// TwinCAT 3 PLC project TcoAteqMeasurement
// Title: TcoAteqMeasurement
// Company: Vortex.Library
// ProjectVersion: 0.6.0.913
// ProgramVersion: 3.1.4023.0
// libraries:
//   Tc2_Standard, * (Beckhoff Automation GmbH)
//   Tc2_System, * (Beckhoff Automation GmbH)
//   Tc3_Module, * (Beckhoff Automation GmbH)
//   TcoIo, 0.6.0.913 (Vortex.Library)
//   TcoCore, 0.6.0.913 (Vortex.Library)
// project tree:
//   DUTs/G6/Enums/ eTcoAteqG6_AlarmCode_v_3_5_x.TcDUT, eTcoAteqG6_ParameterId_v_3_5_x.TcDUT, eTcoAteqG6_SpecialCycle_v_3_5_x.TcDUT, eTcoAteqG6_Step_v_3_5_x.TcDUT, eTcoAteqG6_TestType_v_3_5_x.TcDUT, eTcoAteqG6_Unit_v_3_5_x.TcDUT
//   DUTs/G6/ TcoAteqG6_CommandBits_v_3_5_x.TcDUT, TcoAteqG6_Config_v_3_5_x.TcDUT, TcoAteqG6_Control_v_3_5_x.TcDUT, TcoAteqG6_LastResult_v_3_5_x.TcDUT, TcoAteqG6_Measurement_v_3_5_x.TcDUT, TcoAteqG6_Parameter_v_3_5_x.TcDUT, TcoAteqG6_ParameterList_v_3_5_x.TcDUT, TcoAteqG6_ParameterQuery_v_3_5_x.TcDUT, TcoAteqG6_ParameterRequest_v_3_5_x.TcDUT, TcoAteqG6_ParameterSet_v_3_5_x.TcDUT, TcoAteqG6_State_v_3_5_x.TcDUT, TcoAteqG6_Status_v_3_5_x.TcDUT, TcoAteqG6_StatusBits_v_3_5_x.TcDUT
//   / PlcTask.TcTTO
//   POUs/Functions/G6/ TcoAteqG6_AddParameterToRequest_v_3_5_x.TcPOU, TcoAteqG6_BuildPresetRequest_v_3_5_x.TcPOU, TcoAteqG6_ClearLastResult_v_3_5_x.TcPOU, TcoAteqG6_ClearMeasurement_v_3_5_x.TcPOU, TcoAteqG6_ClearParameterList_v_3_5_x.TcPOU, TcoAteqG6_ClearParameterRequest_v_3_5_x.TcPOU, TcoAteqG6_DecodeCommandBits_v_3_5_x.TcPOU, TcoAteqG6_DecodeLastResult_v_3_5_x.TcPOU, TcoAteqG6_DecodeMeasurement_v_3_5_x.TcPOU, TcoAteqG6_DecodeParameterList_v_3_5_x.TcPOU, TcoAteqG6_DecodeState_v_3_5_x.TcPOU, TcoAteqG6_DecodeStatusBits_v_3_5_x.TcPOU, TcoAteqG6_EncodeControl_v_3_5_x.TcPOU, TcoAteqG6_GetDint_v_3_5_x.TcPOU, TcoAteqG6_GetInt_v_3_5_x.TcPOU, TcoAteqG6_GetWord_v_3_5_x.TcPOU, TcoAteqG6_IsParameterRequestValid_v_3_5_x.TcPOU, TcoAteqG6_MapPresetParameters_v_3_5_x.TcPOU, TcoAteqG6_QueryParameter_v_3_5_x.TcPOU, TcoAteqG6_SetDint_v_3_5_x.TcPOU, TcoAteqG6_SetWord_v_3_5_x.TcPOU, TcoAteqG6_SpecialCycleToByte_v_3_5_x.TcPOU, TcoAteqG6_ToAlarmCode_v_3_5_x.TcPOU, TcoAteqG6_ToEngineering_v_3_5_x.TcPOU, TcoAteqG6_ToStep_v_3_5_x.TcPOU, TcoAteqG6_ToTestType_v_3_5_x.TcPOU, TcoAteqG6_ToUnit_v_3_5_x.TcPOU, TcoAteqG6_TryGetParameterRaw_v_3_5_x.TcPOU
//   POUs/ MAIN.TcPOU
//   POUs/Prototypes/G6/IO/ TcoAteqG6_Inputs_v_3_5_x.TcDUT, TcoAteqG6_Outputs_v_3_5_x.TcDUT, TcoAteqG6Pn_IO_v_3_5_x.TcDUT
//   POUs/Prototypes/G6/ TcoAteqG6Pn_v_3_5_x.TcPOU
//   POUs/Prototypes/MeasurementTasks/G6_v_3_5_x/ TcoAteqG6_ReadLastResultTask_v_3_5_x.TcPOU, TcoAteqG6_ReadParametersTask_v_3_5_x.TcPOU, TcoAteqG6_ResetTask_v_3_5_x.TcPOU, TcoAteqG6_SelectProgramTask_v_3_5_x.TcPOU, TcoAteqG6_SpecialCycleTask_v_3_5_x.TcPOU, TcoAteqG6_StartCycleTask_v_3_5_x.TcPOU, TcoAteqG6Task_v_3_5_x.TcPOU
// real-time tasks:
//   TASK PlcTask: cycle T#10ms, priority 20, ADS port 350
//   TASK PlcTask1: cycle T#10ms, priority 21, ADS port 351

CONFIGURATION TcoAteqMeasurement
    RESOURCE PLC ON TwinCAT3
        TASK PlcTask(INTERVAL := T#10ms, PRIORITY := 20);
        PROGRAM MAIN WITH PlcTask : MAIN;
    END_RESOURCE
END_CONFIGURATION

// ---- DUTs/G6/Enums/eTcoAteqG6_AlarmCode_v_3_5_x.TcDUT
(*~
	<docu>
		<summary>
			Alarm code of the last result (exchange zone 26h). Codes that are not listed decode to Unknown.
		</summary>
	</docu>
~*)
{attribute 'qualified_only'}
{attribute 'strict'}
TYPE eTcoAteqG6_AlarmCode_v_3_5_x :
(
	Unknown := -1,
	NoAlarm := 0,
	PressureSwitchTooHigh := 1,
	PressureSwitchTooLow := 2,
	LargeLeakOnTest := 3,
	LargeLeakOnReference := 4,
	SensorOutOfOrder := 7,
	PressureTooHigh := 43,
	PressureTooLow := 44,
	PiezoSensorOutOfOrder := 45,
	DumpError := 46,
	CalibrationDrift := 47,
	AtmosphericPressureError := 73,
	TemperatureError := 74
) INT;
END_TYPE

// ---- DUTs/G6/Enums/eTcoAteqG6_ParameterId_v_3_5_x.TcDUT
(*~
	<docu>
		<summary>
			Parameter identifiers of the "Read parameters" command (manual pp. 43-46). Every value is exchanged as LONG x1000; times in seconds, levels in the instrument units, selections as code x1000.
		</summary>
	</docu>
~*)
{attribute 'qualified_only'}
{attribute 'strict'}
TYPE eTcoAteqG6_ParameterId_v_3_5_x :
(
	None := 0,
	FillTime := 1,
	StabTime := 2,
	TestTime := 3,
	PreFillTime := 6,
	DumpTime := 9,
	CouplingTimeA := 10,
	CouplingTimeB := 11,
	PartVolume := 20,
	TestType := 21,
	InterCycleTime := 29,
	ResultHoldTime := 48,
	MinFill := 50,
	MaxFill := 51,
	PressureUnit := 53,
	TestFail := 60,
	TestRework := 61,
	RefFail := 62,
	RefRework := 63,
	SetFill := 66,
	DiffAutoResetTime := 80,
	FillMode := 103,
	ExternalDumpType := 110,
	Input7Function := 112,
	Language := 123,
	MaxPreFill := 126,
	FlowUnit := 127,
	CalibrationLeakRate := 128,
	Filter := 148,
	UnitType := 149,
	BarGraphMaxReject := 158,
	VolumeUnit := 161,
	NextProgram := 164,
	PiezoAutoZeroCycles := 165,
	PiezoAutoZeroMinutes := 166,
	DelayExt1 := 249,
	DelayExt2 := 250,
	DelayExt3 := 251,
	DelayExt4 := 252,
	DelayExt5 := 253,
	DelayExt6 := 254,
	DelayInt2 := 255,
	DelayInt1 := 256,
	DelayAux1 := 257,
	DelayAux2 := 258,
	DelayAux3 := 259,
	DelayAux4 := 260,
	TimeExt1 := 261,
	TimeExt2 := 262,
	TimeExt3 := 263,
	TimeExt4 := 264,
	TimeExt5 := 265,
	TimeExt6 := 266,
	TimeInt2 := 267,
	TimeInt1 := 268,
	TimeAux1 := 269,
	TimeAux2 := 270,
	TimeAux3 := 271,
	TimeAux4 := 272,
	PressureFilter := 274,
	CapillaryRange := 281,
	BarCodeFirstChar := 287,
	BarCodeCharCount := 288,
	BarCodeProgram := 289,
	GeneralPressureUnit := 353,
	LinePressureMin := 354,
	DisplayMode := 364,
	Input8Function := 375,
	Input9Function := 376,
	UsbMode := 379,
	SaveOn := 412,
	AccessMode := 413,
	Year := 414,
	Month := 415,
	Day := 416,
	Hour := 417,
	Minute := 418,
	Second := 419,
	LearningCycles := 459,
	LearningInterCycleTime := 460,
	LearningMaxOffset := 461,
	LearningFlowMaster := 462,
	LearningPressureMaster := 463,
	LearningMinVolume := 464,
	LearningMaxVolume := 465,
	LearningOffset := 486
) UINT;
END_TYPE

// ---- DUTs/G6/Enums/eTcoAteqG6_SpecialCycle_v_3_5_x.TcDUT
(*~
	<docu>
		<summary>
			Special cycle table (manual p. 58). Ids 25..31 require the "Service" special-cycle function to be enabled on the instrument.
		</summary>
	</docu>
~*)
{attribute 'qualified_only'}
{attribute 'strict'}
TYPE eTcoAteqG6_SpecialCycle_v_3_5_x :
(
	None := 0,
	AtrLearning := 1,
	CustomUnitLearn := 4,
	CustomUnitCheck := 5,
	PiezoAutoZero := 9,
	RegulatorAdjust := 13,
	CapillaryTemperatureCheck := 25,
	TemperatureCheck := 26,
	AtmPressureCheck := 27,
	P1SensorCheck := 28,
	Flow1Check := 29,
	Flow2Check := 30,
	LinePressureSensorCheck := 31
) INT;
END_TYPE

// ---- DUTs/G6/Enums/eTcoAteqG6_Step_v_3_5_x.TcDUT
(*~
	<docu>
		<summary>
			Current test step (input 0Eh). None = FFFFh on the bus (no cycle running).
		</summary>
	</docu>
~*)
{attribute 'qualified_only'}
{attribute 'strict'}
TYPE eTcoAteqG6_Step_v_3_5_x :
(
	Unknown := -2,
	None := -1,
	PreFill := 0,
	Fill := 1,
	ZeroDiff := 2,
	Stabilization := 3,
	Test := 4,
	Dump := 5
) INT;
END_TYPE

// ---- DUTs/G6/Enums/eTcoAteqG6_TestType_v_3_5_x.TcDUT
(*~
	<docu>
		<summary>
			Test type parameter (id 21).
		</summary>
	</docu>
~*)
{attribute 'qualified_only'}
{attribute 'strict'}
TYPE eTcoAteqG6_TestType_v_3_5_x :
(
	Unknown := -1,
	Invalid := 0,
	Direct := 1,
	Operator := 2
) INT;
END_TYPE

// ---- DUTs/G6/Enums/eTcoAteqG6_Unit_v_3_5_x.TcDUT
(*~
	<docu>
		<summary>
			Unit table (manual p. 48). On the bus a unit is a LONG holding the unit code; the enum value is that code divided by 1000 (14000 = mbar).
		</summary>
	</docu>
~*)
{attribute 'qualified_only'}
{attribute 'strict'}
TYPE eTcoAteqG6_Unit_v_3_5_x :
(
	Unknown := -1,
	cm3_s := 0,
	cm3_min := 1,
	cm3_h := 2,
	Pa := 6,
	bar := 11,
	kPa := 12,
	PSI := 13,
	mbar := 14,
	MPa := 15,
	l_h := 30,
	inch3_s := 46,
	inch3_min := 47,
	inch3_h := 48,
	ft3_h := 49,
	ml_s := 50,
	ml_min := 51,
	ml_h := 52,
	mm3 := 55,
	cm3 := 56,
	ml := 61,
	l := 62,
	inch3 := 63,
	ft3 := 64,
	SCCM := 84,
	Points := 92
) INT;
END_TYPE

// ---- DUTs/G6/TcoAteqG6_CommandBits_v_3_5_x.TcDUT
(*~
	<docu>
		<summary>
			Bit view of a command, echo or error word (bit 0 = Reset ... bit 15 = Read last result).
		</summary>
	</docu>
~*)
TYPE TcoAteqG6_CommandBits_v_3_5_x :
STRUCT
	{attribute addProperty Name "<#Raw#>"}
	Raw : WORD;
	{attribute addProperty Name "<#Reset#>"}
	Reset : BOOL;
	{attribute addProperty Name "<#Start#>"}
	Start : BOOL;
	{attribute addProperty Name "<#Special cycle#>"}
	SpecialCycle : BOOL;
	{attribute addProperty Name "<#Program selection#>"}
	ProgramSelection : BOOL;
	{attribute addProperty Name "<#Read FIFO results#>"}
	ReadFifo : BOOL;
	{attribute addProperty Name "<#Read parameters#>"}
	ReadParameters : BOOL;
	{attribute addProperty Name "<#Write parameters#>"}
	WriteParameters : BOOL;
	{attribute addProperty Name "<#Reset FIFO results#>"}
	ResetFifo : BOOL;
	{attribute addProperty Name "<#Read instrument configuration#>"}
	ReadInstrumentConfiguration : BOOL;
	{attribute addProperty Name "<#Read configuration bits#>"}
	ReadConfigurationBits : BOOL;
	{attribute addProperty Name "<#Read function bits#>"}
	ReadFunctionBits : BOOL;
	{attribute addProperty Name "<#Write configuration bits#>"}
	WriteConfigurationBits : BOOL;
	{attribute addProperty Name "<#Write function bits#>"}
	WriteFunctionBits : BOOL;
	{attribute addProperty Name "<#Read program name#>"}
	ReadProgramName : BOOL;
	{attribute addProperty Name "<#Write program name#>"}
	WriteProgramName : BOOL;
	{attribute addProperty Name "<#Read last result#>"}
	ReadLastResult : BOOL;
END_STRUCT
END_TYPE

// ---- DUTs/G6/TcoAteqG6_Config_v_3_5_x.TcDUT
(*~
	<docu>
		<summary>
			Configuration of TcoAteqG6Pn_v_3_5_x. CommandTimeout / CycleTimeout of 0 fall back to 5 s / 60 s.
		</summary>
	</docu>
~*)
TYPE TcoAteqG6_Config_v_3_5_x :
STRUCT
	{attribute addProperty Name "<#Info time#>"}
	InfoTime : TIME := T#2S;
	{attribute addProperty Name "<#Task timeout (0 = off)#>"}
	ErrorTime : TIME := T#0S;
	{attribute addProperty Name "<#Command handshake timeout (per step)#>"}
	CommandTimeout : TIME := T#5S;
	{attribute addProperty Name "<#Test cycle timeout#>"}
	CycleTimeout : TIME := T#60S;
END_STRUCT
END_TYPE

// ---- DUTs/G6/TcoAteqG6_Control_v_3_5_x.TcDUT
(*~
	<docu>
		<summary>
			Output data: 00h command word, 06h program number (0-based on the bus), 08h special cycle id, 09h special cycle instruction, 20h parameter request. The whole output image is rewritten every cycle.
		</summary>
	</docu>
~*)
TYPE TcoAteqG6_Control_v_3_5_x :
STRUCT
	{attribute addProperty Name "<#Command word#>"}
	Command : WORD;
	{attribute addProperty Name "<#Command bits#>"}
	CommandBits : TcoAteqG6_CommandBits_v_3_5_x;
	{attribute addProperty Name "<#Program number (as displayed, 1-128)#>"}
	ProgramNumber : INT;
	{attribute addProperty Name "<#Special cycle#>"}
	SpecialCycle : eTcoAteqG6_SpecialCycle_v_3_5_x;
	{attribute addProperty Name "<#Special cycle instruction#>"}
	SpecialCycleInstruction : BYTE;
	{attribute addProperty Name "<#Parameter request#>"}
	ParameterRequest : TcoAteqG6_ParameterRequest_v_3_5_x;
	{attribute addProperty Name "<#Selected parameter#>"}
	QueryParameter : eTcoAteqG6_ParameterId_v_3_5_x;
END_STRUCT
END_TYPE

// ---- DUTs/G6/TcoAteqG6_LastResult_v_3_5_x.TcDUT
(*~
	<docu>
		<summary>
			Last result, decoded from the exchange zone (20h..37h) after the "Read last result" command. Valid = no alarm.
		</summary>
	</docu>
~*)
TYPE TcoAteqG6_LastResult_v_3_5_x :
STRUCT
	{attribute addProperty Name "<#Valid#>"}
	Valid : BOOL;
	{attribute addProperty Name "<#Program#>"}
	ProgramNo : INT;
	{attribute addProperty Name "<#Test type (raw)#>"}
	TestTypeRaw : INT;
	{attribute addProperty Name "<#Pass#>"}
	Pass : BOOL;
	{attribute addProperty Name "<#Fail test part (maximum flow reject)#>"}
	FailTest : BOOL;
	{attribute addProperty Name "<#Fail reference part (minimum flow reject)#>"}
	FailReference : BOOL;
	{attribute addProperty Name "<#Alarm#>"}
	Alarm : BOOL;
	{attribute addProperty Name "<#Pressure error (unverified)#>"}
	PressureError : BOOL;
	{attribute addProperty Name "<#Part recoverable (unverified)#>"}
	Recoverable : BOOL;
	{attribute addProperty Name "<#Calibration error (unverified)#>"}
	CalibrationError : BOOL;
	{attribute addProperty Name "<#Calibration check error (unverified)#>"}
	CalibrationCheckError : BOOL;
	{attribute addProperty Name "<#ATR fault (unverified)#>"}
	AtrFault : BOOL;
	{attribute addProperty Name "<#Relay image (raw)#>"}
	RelayImageRaw : WORD;
	{attribute addProperty Name "<#Alarm code#>"}
	AlarmCode : eTcoAteqG6_AlarmCode_v_3_5_x;
	{attribute addProperty Name "<#Alarm code (raw)#>"}
	AlarmCodeRaw : INT;
	{attribute addProperty Name "<#Measurement#>"}
	Measurement : TcoAteqG6_Measurement_v_3_5_x;
END_STRUCT
END_TYPE

// ---- DUTs/G6/TcoAteqG6_Measurement_v_3_5_x.TcDUT
(*~
	<docu>
		<summary>
			Pressure and flow with their units: four LONGs (value x1000, unit code).
		</summary>
	</docu>
~*)
TYPE TcoAteqG6_Measurement_v_3_5_x :
STRUCT
	{attribute addProperty Name "<#Pressure#>"}
	Pressure : REAL;
	{attribute addProperty Name "<#Pressure unit#>"}
	PressureUnit : eTcoAteqG6_Unit_v_3_5_x := eTcoAteqG6_Unit_v_3_5_x.Unknown;
	{attribute addProperty Name "<#Flow / leak#>"}
	Flow : REAL;
	{attribute addProperty Name "<#Flow unit#>"}
	FlowUnit : eTcoAteqG6_Unit_v_3_5_x := eTcoAteqG6_Unit_v_3_5_x.Unknown;
	{attribute addProperty Name "<#Pressure (raw x1000)#>"}
	PressureRaw : DINT;
	{attribute addProperty Name "<#Pressure unit code (raw)#>"}
	PressureUnitRaw : DINT;
	{attribute addProperty Name "<#Flow (raw x1000)#>"}
	FlowRaw : DINT;
	{attribute addProperty Name "<#Flow unit code (raw)#>"}
	FlowUnitRaw : DINT;
END_STRUCT
END_TYPE

// ---- DUTs/G6/TcoAteqG6_Parameter_v_3_5_x.TcDUT
(*~
	<docu>
		<summary>
			One parameter of the "Read parameters" response.
		</summary>
	</docu>
~*)
TYPE TcoAteqG6_Parameter_v_3_5_x :
STRUCT
	{attribute addProperty Name "<#Identifier#>"}
	Id : UINT;
	{attribute addProperty Name "<#Value#>"}
	Value : REAL;
	{attribute addProperty Name "<#Value (raw x1000)#>"}
	Raw : DINT;
END_STRUCT
END_TYPE

// ---- DUTs/G6/TcoAteqG6_ParameterList_v_3_5_x.TcDUT
(*~
	<docu>
		<summary>
			Response of the "Read parameters" command: from input 20h one identifier WORD + value LONG x1000 per parameter.
		</summary>
	</docu>
~*)
TYPE TcoAteqG6_ParameterList_v_3_5_x :
STRUCT
	{attribute addProperty Name "<#Number of parameters read#>"}
	Count : INT;
	{attribute addProperty Name "<#Parameters#>"}
	Items : ARRAY[0..34] OF TcoAteqG6_Parameter_v_3_5_x;
END_STRUCT
END_TYPE

// ---- DUTs/G6/TcoAteqG6_ParameterQuery_v_3_5_x.TcDUT
(*~
	<docu>
		<summary>
			Value of the selected parameter (Control.QueryParameter), looked up after every "Read parameters".
		</summary>
	</docu>
~*)
TYPE TcoAteqG6_ParameterQuery_v_3_5_x :
STRUCT
	{attribute addProperty Name "<#Parameter#>"}
	Parameter : eTcoAteqG6_ParameterId_v_3_5_x;
	{attribute addProperty Name "<#Found#>"}
	Found : BOOL;
	{attribute addProperty Name "<#Value#>"}
	Value : REAL;
	{attribute addProperty Name "<#Value (raw x1000)#>"}
	Raw : DINT;
END_STRUCT
END_TYPE

// ---- DUTs/G6/TcoAteqG6_ParameterRequest_v_3_5_x.TcDUT
(*~
	<docu>
		<summary>
			Request of the "Read parameters" command (output 20h: count, then up to 35 identifiers).
		</summary>
	</docu>
~*)
TYPE TcoAteqG6_ParameterRequest_v_3_5_x :
STRUCT
	{attribute addProperty Name "<#Number of parameters (1-35)#>"}
	Count : INT;
	{attribute addProperty Name "<#Identifiers#>"}
	Ids : ARRAY[0..34] OF UINT;
END_STRUCT
END_TYPE

// ---- DUTs/G6/TcoAteqG6_ParameterSet_v_3_5_x.TcDUT
(*~
	<docu>
		<summary>
			Typed view of the commonly used program parameters (manual p. 43), filled by ReadPresetParameters.
		</summary>
	</docu>
~*)
TYPE TcoAteqG6_ParameterSet_v_3_5_x :
STRUCT
	{attribute addProperty Name "<#Fill time [s]#>"}
	FillTime : REAL;
	{attribute addProperty Name "<#Stabilization time [s]#>"}
	StabTime : REAL;
	{attribute addProperty Name "<#Test time [s]#>"}
	TestTime : REAL;
	{attribute addProperty Name "<#Dump time [s]#>"}
	DumpTime : REAL;
	{attribute addProperty Name "<#Test type#>"}
	TestType : eTcoAteqG6_TestType_v_3_5_x;
	{attribute addProperty Name "<#Minimum fill pressure#>"}
	MinFill : REAL;
	{attribute addProperty Name "<#Maximum fill pressure#>"}
	MaxFill : REAL;
	{attribute addProperty Name "<#Pressure unit#>"}
	PressureUnit : eTcoAteqG6_Unit_v_3_5_x := eTcoAteqG6_Unit_v_3_5_x.Unknown;
	{attribute addProperty Name "<#Test part reject level#>"}
	TestFail : REAL;
	{attribute addProperty Name "<#Reference part reject level#>"}
	RefFail : REAL;
	{attribute addProperty Name "<#Fill set point#>"}
	SetFill : REAL;
END_STRUCT
END_TYPE

// ---- DUTs/G6/TcoAteqG6_State_v_3_5_x.TcDUT
(*~
	<docu>
		<summary>
			Decoded input image: 00h echo, 02h error word (FFFFh = command running), 06h program (0-based on the bus), 08h results in FIFO, 0Ah test type, 0Ch status bits, 0Eh step, 10h..1Fh real-time pressure/flow.
		</summary>
	</docu>
~*)
TYPE TcoAteqG6_State_v_3_5_x :
STRUCT
	{attribute addProperty Name "<#Command echo#>"}
	Echo : TcoAteqG6_CommandBits_v_3_5_x;
	{attribute addProperty Name "<#Command error#>"}
	Error : TcoAteqG6_CommandBits_v_3_5_x;
	{attribute addProperty Name "<#Command running#>"}
	CommandRunning : BOOL;
	{attribute addProperty Name "<#Current program#>"}
	CurrentProgram : INT;
	{attribute addProperty Name "<#Results in FIFO#>"}
	ResultsInFifo : INT;
	{attribute addProperty Name "<#Test type (raw)#>"}
	TestTypeRaw : INT;
	{attribute addProperty Name "<#Status#>"}
	StatusBits : TcoAteqG6_StatusBits_v_3_5_x;
	{attribute addProperty Name "<#Step#>"}
	Step : eTcoAteqG6_Step_v_3_5_x := eTcoAteqG6_Step_v_3_5_x.None;
	{attribute addProperty Name "<#Step (raw)#>"}
	StepRaw : INT;
	{attribute addProperty Name "<#Real time#>"}
	RealTime : TcoAteqG6_Measurement_v_3_5_x;
END_STRUCT
END_TYPE

// ---- DUTs/G6/TcoAteqG6_Status_v_3_5_x.TcDUT
(*~
	<docu>
		<summary>
			Status of TcoAteqG6Pn_v_3_5_x.
		</summary>
	</docu>
~*)
TYPE TcoAteqG6_Status_v_3_5_x :
STRUCT
	{attribute addProperty Name "<#Action#>"}
	ActionDescription : STRING(100);
	{attribute addProperty Name "<#Ready#>"}
	Ready : BOOL;
	{attribute addProperty Name "<#Last part passed#>"}
	LastPass : BOOL;
	{attribute addProperty Name "<#Last command error word#>"}
	LastCommandError : WORD;
	{attribute addProperty Name "<#Instrument#>"}
	State : TcoAteqG6_State_v_3_5_x;
	{attribute addProperty Name "<#Last result#>"}
	LastResult : TcoAteqG6_LastResult_v_3_5_x;
	{attribute addProperty Name "<#Parameters#>"}
	Parameters : TcoAteqG6_ParameterList_v_3_5_x;
	{attribute addProperty Name "<#Preset parameters#>"}
	ParameterSet : TcoAteqG6_ParameterSet_v_3_5_x;
	{attribute addProperty Name "<#Selected parameter#>"}
	ParameterQuery : TcoAteqG6_ParameterQuery_v_3_5_x;
END_STRUCT
END_TYPE

// ---- DUTs/G6/TcoAteqG6_StatusBits_v_3_5_x.TcDUT
(*~
	<docu>
		<summary>
			Status word of the instrument (input 0Ch). Bits 8 and 10..14 are not used.
		</summary>
	</docu>
~*)
TYPE TcoAteqG6_StatusBits_v_3_5_x :
STRUCT
	{attribute addProperty Name "<#Raw#>"}
	Raw : WORD;
	{attribute addProperty Name "<#Pass#>"}
	Pass : BOOL;
	{attribute addProperty Name "<#Fail test part#>"}
	FailTest : BOOL;
	{attribute addProperty Name "<#Fail reference part#>"}
	FailReference : BOOL;
	{attribute addProperty Name "<#Alarm#>"}
	Alarm : BOOL;
	{attribute addProperty Name "<#Pressure error#>"}
	PressureError : BOOL;
	{attribute addProperty Name "<#Cycle end#>"}
	CycleEnd : BOOL;
	{attribute addProperty Name "<#Part recoverable#>"}
	Recoverable : BOOL;
	{attribute addProperty Name "<#Calibration error or drift#>"}
	CalibrationError : BOOL;
	{attribute addProperty Name "<#ATR error or drift#>"}
	AtrError : BOOL;
	{attribute addProperty Name "<#Key presence#>"}
	KeyPresence : BOOL;
END_STRUCT
END_TYPE

// ---- POUs/Prototypes/G6/IO/TcoAteqG6_Inputs_v_3_5_x.TcDUT
TYPE TcoAteqG6_Inputs_v_3_5_x :
STRUCT
	{attribute addProperty Name "<#Input module 1 (slot 1, 00h..3Fh)#>"}
	In1 AT %I* : ARRAY[0..63] OF BYTE;
	{attribute addProperty Name "<#Input module 2 (slot 2, 40h..7Fh)#>"}
	In2 AT %I* : ARRAY[0..63] OF BYTE;
	{attribute addProperty Name "<#Input module 3 (slot 3, 80h..BFh)#>"}
	In3 AT %I* : ARRAY[0..63] OF BYTE;
	{attribute addProperty Name "<#Input module 4 (slot 4, C0h..FFh)#>"}
	In4 AT %I* : ARRAY[0..63] OF BYTE;
END_STRUCT
END_TYPE

// ---- POUs/Prototypes/G6/IO/TcoAteqG6_Outputs_v_3_5_x.TcDUT
TYPE TcoAteqG6_Outputs_v_3_5_x :
STRUCT
	{attribute addProperty Name "<#Output module 1 (slot 5, 00h..3Fh)#>"}
	Out1 AT %Q* : ARRAY[0..63] OF BYTE;
	{attribute addProperty Name "<#Output module 2 (slot 6, 40h..7Fh)#>"}
	Out2 AT %Q* : ARRAY[0..63] OF BYTE;
	{attribute addProperty Name "<#Output module 3 (slot 7, 80h..BFh)#>"}
	Out3 AT %Q* : ARRAY[0..63] OF BYTE;
	{attribute addProperty Name "<#Output module 4 (slot 8, C0h..FFh)#>"}
	Out4 AT %Q* : ARRAY[0..63] OF BYTE;
END_STRUCT
END_TYPE

// ---- POUs/Prototypes/G6/IO/TcoAteqG6Pn_IO_v_3_5_x.TcDUT
TYPE TcoAteqG6Pn_IO_v_3_5_x :
STRUCT
	PnIoBoxState AT %I*	:	UINT;
	PnIoBoxDiag AT %I*	:	UINT;
	PnIoBoxCtrl AT %Q*	:	UINT;
	{attribute addProperty Name "<#IN#>"}
	In : TcoAteqG6_Inputs_v_3_5_x;
	{attribute addProperty Name "<#OUT#>"}
	Out : TcoAteqG6_Outputs_v_3_5_x;
END_STRUCT
END_TYPE

// ---- POUs/MAIN.TcPOU
PROGRAM MAIN
VAR
END_VAR

END_PROGRAM

// ---- POUs/Functions/G6/TcoAteqG6_AddParameterToRequest_v_3_5_x.TcPOU
(*~
	<docu>
		<summary>
			Appends a parameter identifier to the request. Returns FALSE when the request is full (35).
		</summary>
	</docu>
~*)
FUNCTION TcoAteqG6_AddParameterToRequest_v_3_5_x : BOOL
VAR_INPUT
	inParameter : eTcoAteqG6_ParameterId_v_3_5_x;
END_VAR
VAR_IN_OUT
	inoRequest : TcoAteqG6_ParameterRequest_v_3_5_x;
END_VAR

IF inoRequest.Count < 0 OR inoRequest.Count >= 35 THEN
	RETURN;
END_IF
inoRequest.Ids[inoRequest.Count] := TO_UINT(inParameter);
inoRequest.Count := inoRequest.Count + 1;
TcoAteqG6_AddParameterToRequest_v_3_5_x := TRUE;

END_FUNCTION

// ---- POUs/Functions/G6/TcoAteqG6_BuildPresetRequest_v_3_5_x.TcPOU
(*~
	<docu>
		<summary>
			Fills the request with the 11 identifiers of the preset parameter set.
		</summary>
	</docu>
~*)
FUNCTION TcoAteqG6_BuildPresetRequest_v_3_5_x : BOOL
VAR_IN_OUT
	inoRequest : TcoAteqG6_ParameterRequest_v_3_5_x;
END_VAR

TcoAteqG6_ClearParameterRequest_v_3_5_x(inoRequest := inoRequest);
TcoAteqG6_AddParameterToRequest_v_3_5_x(inParameter := eTcoAteqG6_ParameterId_v_3_5_x.FillTime, inoRequest := inoRequest);
TcoAteqG6_AddParameterToRequest_v_3_5_x(inParameter := eTcoAteqG6_ParameterId_v_3_5_x.StabTime, inoRequest := inoRequest);
TcoAteqG6_AddParameterToRequest_v_3_5_x(inParameter := eTcoAteqG6_ParameterId_v_3_5_x.TestTime, inoRequest := inoRequest);
TcoAteqG6_AddParameterToRequest_v_3_5_x(inParameter := eTcoAteqG6_ParameterId_v_3_5_x.DumpTime, inoRequest := inoRequest);
TcoAteqG6_AddParameterToRequest_v_3_5_x(inParameter := eTcoAteqG6_ParameterId_v_3_5_x.TestType, inoRequest := inoRequest);
TcoAteqG6_AddParameterToRequest_v_3_5_x(inParameter := eTcoAteqG6_ParameterId_v_3_5_x.MinFill, inoRequest := inoRequest);
TcoAteqG6_AddParameterToRequest_v_3_5_x(inParameter := eTcoAteqG6_ParameterId_v_3_5_x.MaxFill, inoRequest := inoRequest);
TcoAteqG6_AddParameterToRequest_v_3_5_x(inParameter := eTcoAteqG6_ParameterId_v_3_5_x.PressureUnit, inoRequest := inoRequest);
TcoAteqG6_AddParameterToRequest_v_3_5_x(inParameter := eTcoAteqG6_ParameterId_v_3_5_x.TestFail, inoRequest := inoRequest);
TcoAteqG6_AddParameterToRequest_v_3_5_x(inParameter := eTcoAteqG6_ParameterId_v_3_5_x.RefFail, inoRequest := inoRequest);
TcoAteqG6_AddParameterToRequest_v_3_5_x(inParameter := eTcoAteqG6_ParameterId_v_3_5_x.SetFill, inoRequest := inoRequest);
TcoAteqG6_BuildPresetRequest_v_3_5_x := TRUE;

END_FUNCTION

// ---- POUs/Functions/G6/TcoAteqG6_ClearParameterRequest_v_3_5_x.TcPOU
(*~
	<docu>
		<summary>
			Clears a parameter request.
		</summary>
	</docu>
~*)
FUNCTION TcoAteqG6_ClearParameterRequest_v_3_5_x : BOOL
VAR_IN_OUT
	inoRequest : TcoAteqG6_ParameterRequest_v_3_5_x;
END_VAR
VAR
	i : INT;
END_VAR

inoRequest.Count := 0;
FOR i := 0 TO 34 DO
	inoRequest.Ids[i] := 0;
END_FOR
TcoAteqG6_ClearParameterRequest_v_3_5_x := TRUE;

END_FUNCTION

// ---- POUs/Functions/G6/TcoAteqG6_ClearLastResult_v_3_5_x.TcPOU
(*~
	<docu>
		<summary>
			Clears the last result (Valid = FALSE).
		</summary>
	</docu>
~*)
FUNCTION TcoAteqG6_ClearLastResult_v_3_5_x : BOOL
VAR_IN_OUT
	inoResult : TcoAteqG6_LastResult_v_3_5_x;
END_VAR

inoResult.Valid := FALSE;
inoResult.ProgramNo := 0;
inoResult.TestTypeRaw := 0;
inoResult.Pass := FALSE;
inoResult.FailTest := FALSE;
inoResult.FailReference := FALSE;
inoResult.Alarm := FALSE;
inoResult.PressureError := FALSE;
inoResult.Recoverable := FALSE;
inoResult.CalibrationError := FALSE;
inoResult.CalibrationCheckError := FALSE;
inoResult.AtrFault := FALSE;
inoResult.RelayImageRaw := 0;
inoResult.AlarmCode := eTcoAteqG6_AlarmCode_v_3_5_x.NoAlarm;
inoResult.AlarmCodeRaw := 0;
TcoAteqG6_ClearMeasurement_v_3_5_x(inoMeasurement := inoResult.Measurement);
TcoAteqG6_ClearLastResult_v_3_5_x := TRUE;

END_FUNCTION

// ---- POUs/Functions/G6/TcoAteqG6_ClearMeasurement_v_3_5_x.TcPOU
(*~
	<docu>
		<summary>
			Clears a measurement.
		</summary>
	</docu>
~*)
FUNCTION TcoAteqG6_ClearMeasurement_v_3_5_x : BOOL
VAR_IN_OUT
	inoMeasurement : TcoAteqG6_Measurement_v_3_5_x;
END_VAR

inoMeasurement.Pressure := 0.0;
inoMeasurement.PressureUnit := eTcoAteqG6_Unit_v_3_5_x.Unknown;
inoMeasurement.Flow := 0.0;
inoMeasurement.FlowUnit := eTcoAteqG6_Unit_v_3_5_x.Unknown;
inoMeasurement.PressureRaw := 0;
inoMeasurement.PressureUnitRaw := 0;
inoMeasurement.FlowRaw := 0;
inoMeasurement.FlowUnitRaw := 0;
TcoAteqG6_ClearMeasurement_v_3_5_x := TRUE;

END_FUNCTION

// ---- POUs/Functions/G6/TcoAteqG6_ClearParameterList_v_3_5_x.TcPOU
(*~
	<docu>
		<summary>
			Clears a parameter list.
		</summary>
	</docu>
~*)
FUNCTION TcoAteqG6_ClearParameterList_v_3_5_x : BOOL
VAR_IN_OUT
	inoList : TcoAteqG6_ParameterList_v_3_5_x;
END_VAR
VAR
	i : INT;
END_VAR

inoList.Count := 0;
FOR i := 0 TO 34 DO
	inoList.Items[i].Id := 0;
	inoList.Items[i].Raw := 0;
	inoList.Items[i].Value := 0.0;
END_FOR
TcoAteqG6_ClearParameterList_v_3_5_x := TRUE;

END_FUNCTION

// ---- POUs/Functions/G6/TcoAteqG6_DecodeCommandBits_v_3_5_x.TcPOU
(*~
	<docu>
		<summary>
			Bit view of a command, echo or error word.
		</summary>
	</docu>
~*)
FUNCTION TcoAteqG6_DecodeCommandBits_v_3_5_x : BOOL
VAR_INPUT
	inValue : WORD;
END_VAR
VAR_IN_OUT
	inoBits : TcoAteqG6_CommandBits_v_3_5_x;
END_VAR

inoBits.Raw := inValue;
inoBits.Reset := inValue.0;
inoBits.Start := inValue.1;
inoBits.SpecialCycle := inValue.2;
inoBits.ProgramSelection := inValue.3;
inoBits.ReadFifo := inValue.4;
inoBits.ReadParameters := inValue.5;
inoBits.WriteParameters := inValue.6;
inoBits.ResetFifo := inValue.7;
inoBits.ReadInstrumentConfiguration := inValue.8;
inoBits.ReadConfigurationBits := inValue.9;
inoBits.ReadFunctionBits := inValue.10;
inoBits.WriteConfigurationBits := inValue.11;
inoBits.WriteFunctionBits := inValue.12;
inoBits.ReadProgramName := inValue.13;
inoBits.WriteProgramName := inValue.14;
inoBits.ReadLastResult := inValue.15;
TcoAteqG6_DecodeCommandBits_v_3_5_x := TRUE;

END_FUNCTION

// ---- POUs/Functions/G6/TcoAteqG6_DecodeLastResult_v_3_5_x.TcPOU
(*~
	<docu>
		<summary>
			Decodes the last result from the exchange zone (20h program, 22h test type, 24h relay image, 26h alarm code, 28h..37h measurement). Relay bits 4..8 are not verified on hardware.
		</summary>
	</docu>
~*)
FUNCTION TcoAteqG6_DecodeLastResult_v_3_5_x : BOOL
VAR_IN_OUT
	inoImage : ARRAY[0..255] OF BYTE;
	inoResult : TcoAteqG6_LastResult_v_3_5_x;
END_VAR

inoResult.ProgramNo := TcoAteqG6_GetInt_v_3_5_x(inOffset := 16#20, inoImage := inoImage) + 1;
inoResult.TestTypeRaw := TcoAteqG6_GetInt_v_3_5_x(inOffset := 16#22, inoImage := inoImage);
inoResult.RelayImageRaw := TcoAteqG6_GetWord_v_3_5_x(inOffset := 16#24, inoImage := inoImage);
inoResult.Pass := inoResult.RelayImageRaw.0;
inoResult.FailTest := inoResult.RelayImageRaw.1;
inoResult.FailReference := inoResult.RelayImageRaw.2;
inoResult.Alarm := inoResult.RelayImageRaw.3;
inoResult.PressureError := inoResult.RelayImageRaw.4;
inoResult.Recoverable := inoResult.RelayImageRaw.5;
inoResult.CalibrationError := inoResult.RelayImageRaw.6;
inoResult.CalibrationCheckError := inoResult.RelayImageRaw.7;
inoResult.AtrFault := inoResult.RelayImageRaw.8;
inoResult.AlarmCodeRaw := TcoAteqG6_GetInt_v_3_5_x(inOffset := 16#26, inoImage := inoImage);
inoResult.AlarmCode := TcoAteqG6_ToAlarmCode_v_3_5_x(inoResult.AlarmCodeRaw);
TcoAteqG6_DecodeMeasurement_v_3_5_x(inOffset := 16#28, inoImage := inoImage, inoMeasurement := inoResult.Measurement);
inoResult.Valid := NOT inoResult.Alarm;
TcoAteqG6_DecodeLastResult_v_3_5_x := TRUE;

END_FUNCTION

// ---- POUs/Functions/G6/TcoAteqG6_GetInt_v_3_5_x.TcPOU
(*~
	<docu>
		<summary>
			Little-endian INT at inOffset.
		</summary>
	</docu>
~*)
FUNCTION TcoAteqG6_GetInt_v_3_5_x : INT
VAR_INPUT
	inOffset : INT;
END_VAR
VAR_IN_OUT
	inoImage : ARRAY[0..255] OF BYTE;
END_VAR

TcoAteqG6_GetInt_v_3_5_x := WORD_TO_INT(TcoAteqG6_GetWord_v_3_5_x(inOffset := inOffset, inoImage := inoImage));

END_FUNCTION

// ---- POUs/Functions/G6/TcoAteqG6_GetWord_v_3_5_x.TcPOU
(*~
	<docu>
		<summary>
			Little-endian WORD at inOffset (ATEQ fieldbus data: least significant byte first).
		</summary>
	</docu>
~*)
FUNCTION TcoAteqG6_GetWord_v_3_5_x : WORD
VAR_INPUT
	inOffset : INT;
END_VAR
VAR_IN_OUT
	inoImage : ARRAY[0..255] OF BYTE;
END_VAR

TcoAteqG6_GetWord_v_3_5_x := SHL(BYTE_TO_WORD(inoImage[inOffset + 1]), 8) OR BYTE_TO_WORD(inoImage[inOffset]);

END_FUNCTION

// ---- POUs/Functions/G6/TcoAteqG6_ToAlarmCode_v_3_5_x.TcPOU
(*~
	<docu>
		<summary>
			Alarm code word to alarm code.
		</summary>
	</docu>
~*)
FUNCTION TcoAteqG6_ToAlarmCode_v_3_5_x : eTcoAteqG6_AlarmCode_v_3_5_x
VAR_INPUT
	inRaw : INT;
END_VAR

CASE inRaw OF
	0: TcoAteqG6_ToAlarmCode_v_3_5_x := eTcoAteqG6_AlarmCode_v_3_5_x.NoAlarm;
	1: TcoAteqG6_ToAlarmCode_v_3_5_x := eTcoAteqG6_AlarmCode_v_3_5_x.PressureSwitchTooHigh;
	2: TcoAteqG6_ToAlarmCode_v_3_5_x := eTcoAteqG6_AlarmCode_v_3_5_x.PressureSwitchTooLow;
	3: TcoAteqG6_ToAlarmCode_v_3_5_x := eTcoAteqG6_AlarmCode_v_3_5_x.LargeLeakOnTest;
	4: TcoAteqG6_ToAlarmCode_v_3_5_x := eTcoAteqG6_AlarmCode_v_3_5_x.LargeLeakOnReference;
	7: TcoAteqG6_ToAlarmCode_v_3_5_x := eTcoAteqG6_AlarmCode_v_3_5_x.SensorOutOfOrder;
	43: TcoAteqG6_ToAlarmCode_v_3_5_x := eTcoAteqG6_AlarmCode_v_3_5_x.PressureTooHigh;
	44: TcoAteqG6_ToAlarmCode_v_3_5_x := eTcoAteqG6_AlarmCode_v_3_5_x.PressureTooLow;
	45: TcoAteqG6_ToAlarmCode_v_3_5_x := eTcoAteqG6_AlarmCode_v_3_5_x.PiezoSensorOutOfOrder;
	46: TcoAteqG6_ToAlarmCode_v_3_5_x := eTcoAteqG6_AlarmCode_v_3_5_x.DumpError;
	47: TcoAteqG6_ToAlarmCode_v_3_5_x := eTcoAteqG6_AlarmCode_v_3_5_x.CalibrationDrift;
	73: TcoAteqG6_ToAlarmCode_v_3_5_x := eTcoAteqG6_AlarmCode_v_3_5_x.AtmosphericPressureError;
	74: TcoAteqG6_ToAlarmCode_v_3_5_x := eTcoAteqG6_AlarmCode_v_3_5_x.TemperatureError;
ELSE
	TcoAteqG6_ToAlarmCode_v_3_5_x := eTcoAteqG6_AlarmCode_v_3_5_x.Unknown;
END_CASE

END_FUNCTION

// ---- POUs/Functions/G6/TcoAteqG6_DecodeMeasurement_v_3_5_x.TcPOU
(*~
	<docu>
		<summary>
			Decodes pressure, pressure unit, flow and flow unit (4 LONGs) from inOffset.
		</summary>
	</docu>
~*)
FUNCTION TcoAteqG6_DecodeMeasurement_v_3_5_x : BOOL
VAR_INPUT
	inOffset : INT;
END_VAR
VAR_IN_OUT
	inoImage : ARRAY[0..255] OF BYTE;
	inoMeasurement : TcoAteqG6_Measurement_v_3_5_x;
END_VAR

inoMeasurement.PressureRaw := TcoAteqG6_GetDint_v_3_5_x(inOffset := inOffset, inoImage := inoImage);
inoMeasurement.PressureUnitRaw := TcoAteqG6_GetDint_v_3_5_x(inOffset := inOffset + 4, inoImage := inoImage);
inoMeasurement.FlowRaw := TcoAteqG6_GetDint_v_3_5_x(inOffset := inOffset + 8, inoImage := inoImage);
inoMeasurement.FlowUnitRaw := TcoAteqG6_GetDint_v_3_5_x(inOffset := inOffset + 12, inoImage := inoImage);
inoMeasurement.Pressure := TcoAteqG6_ToEngineering_v_3_5_x(inoMeasurement.PressureRaw);
inoMeasurement.PressureUnit := TcoAteqG6_ToUnit_v_3_5_x(inoMeasurement.PressureUnitRaw);
inoMeasurement.Flow := TcoAteqG6_ToEngineering_v_3_5_x(inoMeasurement.FlowRaw);
inoMeasurement.FlowUnit := TcoAteqG6_ToUnit_v_3_5_x(inoMeasurement.FlowUnitRaw);
TcoAteqG6_DecodeMeasurement_v_3_5_x := TRUE;

END_FUNCTION

// ---- POUs/Functions/G6/TcoAteqG6_GetDint_v_3_5_x.TcPOU
(*~
	<docu>
		<summary>
			Little-endian LONG at inOffset (least significant word first).
		</summary>
	</docu>
~*)
FUNCTION TcoAteqG6_GetDint_v_3_5_x : DINT
VAR_INPUT
	inOffset : INT;
END_VAR
VAR_IN_OUT
	inoImage : ARRAY[0..255] OF BYTE;
END_VAR

TcoAteqG6_GetDint_v_3_5_x := DWORD_TO_DINT(SHL(BYTE_TO_DWORD(inoImage[inOffset + 3]), 24)
	OR SHL(BYTE_TO_DWORD(inoImage[inOffset + 2]), 16)
	OR SHL(BYTE_TO_DWORD(inoImage[inOffset + 1]), 8)
	OR BYTE_TO_DWORD(inoImage[inOffset]));

END_FUNCTION

// ---- POUs/Functions/G6/TcoAteqG6_ToEngineering_v_3_5_x.TcPOU
(*~
	<docu>
		<summary>
			Fixed-point LONG (x1000) to engineering value.
		</summary>
	</docu>
~*)
FUNCTION TcoAteqG6_ToEngineering_v_3_5_x : REAL
VAR_INPUT
	inRaw : DINT;
END_VAR

TcoAteqG6_ToEngineering_v_3_5_x := DINT_TO_REAL(inRaw) / 1000.0;

END_FUNCTION

// ---- POUs/Functions/G6/TcoAteqG6_ToUnit_v_3_5_x.TcPOU
(*~
	<docu>
		<summary>
			Unit code (LONG, code x1000) to unit. Codes that are not listed or not a multiple of 1000 give Unknown.
		</summary>
	</docu>
~*)
FUNCTION TcoAteqG6_ToUnit_v_3_5_x : eTcoAteqG6_Unit_v_3_5_x
VAR_INPUT
	inRaw : DINT;
END_VAR
VAR
	code : DINT;
END_VAR

TcoAteqG6_ToUnit_v_3_5_x := eTcoAteqG6_Unit_v_3_5_x.Unknown;
IF inRaw < 0 OR (inRaw MOD 1000) <> 0 THEN
	RETURN;
END_IF
code := inRaw / 1000;
CASE code OF
	0: TcoAteqG6_ToUnit_v_3_5_x := eTcoAteqG6_Unit_v_3_5_x.cm3_s;
	1: TcoAteqG6_ToUnit_v_3_5_x := eTcoAteqG6_Unit_v_3_5_x.cm3_min;
	2: TcoAteqG6_ToUnit_v_3_5_x := eTcoAteqG6_Unit_v_3_5_x.cm3_h;
	6: TcoAteqG6_ToUnit_v_3_5_x := eTcoAteqG6_Unit_v_3_5_x.Pa;
	11: TcoAteqG6_ToUnit_v_3_5_x := eTcoAteqG6_Unit_v_3_5_x.bar;
	12: TcoAteqG6_ToUnit_v_3_5_x := eTcoAteqG6_Unit_v_3_5_x.kPa;
	13: TcoAteqG6_ToUnit_v_3_5_x := eTcoAteqG6_Unit_v_3_5_x.PSI;
	14: TcoAteqG6_ToUnit_v_3_5_x := eTcoAteqG6_Unit_v_3_5_x.mbar;
	15: TcoAteqG6_ToUnit_v_3_5_x := eTcoAteqG6_Unit_v_3_5_x.MPa;
	30: TcoAteqG6_ToUnit_v_3_5_x := eTcoAteqG6_Unit_v_3_5_x.l_h;
	46: TcoAteqG6_ToUnit_v_3_5_x := eTcoAteqG6_Unit_v_3_5_x.inch3_s;
	47: TcoAteqG6_ToUnit_v_3_5_x := eTcoAteqG6_Unit_v_3_5_x.inch3_min;
	48: TcoAteqG6_ToUnit_v_3_5_x := eTcoAteqG6_Unit_v_3_5_x.inch3_h;
	49: TcoAteqG6_ToUnit_v_3_5_x := eTcoAteqG6_Unit_v_3_5_x.ft3_h;
	50: TcoAteqG6_ToUnit_v_3_5_x := eTcoAteqG6_Unit_v_3_5_x.ml_s;
	51: TcoAteqG6_ToUnit_v_3_5_x := eTcoAteqG6_Unit_v_3_5_x.ml_min;
	52: TcoAteqG6_ToUnit_v_3_5_x := eTcoAteqG6_Unit_v_3_5_x.ml_h;
	55: TcoAteqG6_ToUnit_v_3_5_x := eTcoAteqG6_Unit_v_3_5_x.mm3;
	56: TcoAteqG6_ToUnit_v_3_5_x := eTcoAteqG6_Unit_v_3_5_x.cm3;
	61: TcoAteqG6_ToUnit_v_3_5_x := eTcoAteqG6_Unit_v_3_5_x.ml;
	62: TcoAteqG6_ToUnit_v_3_5_x := eTcoAteqG6_Unit_v_3_5_x.l;
	63: TcoAteqG6_ToUnit_v_3_5_x := eTcoAteqG6_Unit_v_3_5_x.inch3;
	64: TcoAteqG6_ToUnit_v_3_5_x := eTcoAteqG6_Unit_v_3_5_x.ft3;
	84: TcoAteqG6_ToUnit_v_3_5_x := eTcoAteqG6_Unit_v_3_5_x.SCCM;
	92: TcoAteqG6_ToUnit_v_3_5_x := eTcoAteqG6_Unit_v_3_5_x.Points;
END_CASE

END_FUNCTION

// ---- POUs/Functions/G6/TcoAteqG6_DecodeParameterList_v_3_5_x.TcPOU
(*~
	<docu>
		<summary>
			Decodes inCount parameters (identifier WORD + value LONG x1000 each) from inOffset. A count outside 1..35 leaves the list empty.
		</summary>
	</docu>
~*)
FUNCTION TcoAteqG6_DecodeParameterList_v_3_5_x : BOOL
VAR_INPUT
	inOffset : INT;
	inCount : INT;
END_VAR
VAR_IN_OUT
	inoImage : ARRAY[0..255] OF BYTE;
	inoList : TcoAteqG6_ParameterList_v_3_5_x;
END_VAR
VAR
	i : INT;
	pos : INT;
END_VAR

TcoAteqG6_ClearParameterList_v_3_5_x(inoList := inoList);
IF inCount < 1 OR inCount > 35 THEN
	RETURN;
END_IF
FOR i := 0 TO inCount - 1 DO
	pos := inOffset + 6 * i;
	inoList.Items[i].Id := WORD_TO_UINT(TcoAteqG6_GetWord_v_3_5_x(inOffset := pos, inoImage := inoImage));
	inoList.Items[i].Raw := TcoAteqG6_GetDint_v_3_5_x(inOffset := pos + 2, inoImage := inoImage);
	inoList.Items[i].Value := TcoAteqG6_ToEngineering_v_3_5_x(inoList.Items[i].Raw);
END_FOR
inoList.Count := inCount;
TcoAteqG6_DecodeParameterList_v_3_5_x := TRUE;

END_FUNCTION

// ---- POUs/Functions/G6/TcoAteqG6_DecodeState_v_3_5_x.TcPOU
(*~
	<docu>
		<summary>
			Decodes the live part of the input image (00h..1Fh). The program number is 0-based on the bus and 1-based here.
		</summary>
	</docu>
~*)
FUNCTION TcoAteqG6_DecodeState_v_3_5_x : BOOL
VAR_IN_OUT
	inoImage : ARRAY[0..255] OF BYTE;
	inoState : TcoAteqG6_State_v_3_5_x;
END_VAR

TcoAteqG6_DecodeCommandBits_v_3_5_x(inValue := TcoAteqG6_GetWord_v_3_5_x(inOffset := 16#00, inoImage := inoImage), inoBits := inoState.Echo);
TcoAteqG6_DecodeCommandBits_v_3_5_x(inValue := TcoAteqG6_GetWord_v_3_5_x(inOffset := 16#02, inoImage := inoImage), inoBits := inoState.Error);
inoState.CommandRunning := inoState.Error.Raw = 16#FFFF;
inoState.CurrentProgram := TcoAteqG6_GetInt_v_3_5_x(inOffset := 16#06, inoImage := inoImage) + 1;
inoState.ResultsInFifo := TcoAteqG6_GetInt_v_3_5_x(inOffset := 16#08, inoImage := inoImage);
inoState.TestTypeRaw := TcoAteqG6_GetInt_v_3_5_x(inOffset := 16#0A, inoImage := inoImage);
TcoAteqG6_DecodeStatusBits_v_3_5_x(inValue := TcoAteqG6_GetWord_v_3_5_x(inOffset := 16#0C, inoImage := inoImage), inoBits := inoState.StatusBits);
inoState.StepRaw := TcoAteqG6_GetInt_v_3_5_x(inOffset := 16#0E, inoImage := inoImage);
inoState.Step := TcoAteqG6_ToStep_v_3_5_x(inoState.StepRaw);
TcoAteqG6_DecodeMeasurement_v_3_5_x(inOffset := 16#10, inoImage := inoImage, inoMeasurement := inoState.RealTime);
TcoAteqG6_DecodeState_v_3_5_x := TRUE;

END_FUNCTION

// ---- POUs/Functions/G6/TcoAteqG6_DecodeStatusBits_v_3_5_x.TcPOU
(*~
	<docu>
		<summary>
			Bit view of the status word (input 0Ch).
		</summary>
	</docu>
~*)
FUNCTION TcoAteqG6_DecodeStatusBits_v_3_5_x : BOOL
VAR_INPUT
	inValue : WORD;
END_VAR
VAR_IN_OUT
	inoBits : TcoAteqG6_StatusBits_v_3_5_x;
END_VAR

inoBits.Raw := inValue;
inoBits.Pass := inValue.0;
inoBits.FailTest := inValue.1;
inoBits.FailReference := inValue.2;
inoBits.Alarm := inValue.3;
inoBits.PressureError := inValue.4;
inoBits.CycleEnd := inValue.5;
inoBits.Recoverable := inValue.6;
inoBits.CalibrationError := inValue.7;
inoBits.AtrError := inValue.9;
inoBits.KeyPresence := inValue.15;
TcoAteqG6_DecodeStatusBits_v_3_5_x := TRUE;

END_FUNCTION

// ---- POUs/Functions/G6/TcoAteqG6_ToStep_v_3_5_x.TcPOU
(*~
	<docu>
		<summary>
			Step word to step.
		</summary>
	</docu>
~*)
FUNCTION TcoAteqG6_ToStep_v_3_5_x : eTcoAteqG6_Step_v_3_5_x
VAR_INPUT
	inRaw : INT;
END_VAR

CASE inRaw OF
	-1: TcoAteqG6_ToStep_v_3_5_x := eTcoAteqG6_Step_v_3_5_x.None;
	0: TcoAteqG6_ToStep_v_3_5_x := eTcoAteqG6_Step_v_3_5_x.PreFill;
	1: TcoAteqG6_ToStep_v_3_5_x := eTcoAteqG6_Step_v_3_5_x.Fill;
	2: TcoAteqG6_ToStep_v_3_5_x := eTcoAteqG6_Step_v_3_5_x.ZeroDiff;
	3: TcoAteqG6_ToStep_v_3_5_x := eTcoAteqG6_Step_v_3_5_x.Stabilization;
	4: TcoAteqG6_ToStep_v_3_5_x := eTcoAteqG6_Step_v_3_5_x.Test;
	5: TcoAteqG6_ToStep_v_3_5_x := eTcoAteqG6_Step_v_3_5_x.Dump;
ELSE
	TcoAteqG6_ToStep_v_3_5_x := eTcoAteqG6_Step_v_3_5_x.Unknown;
END_CASE

END_FUNCTION

// ---- POUs/Functions/G6/TcoAteqG6_EncodeControl_v_3_5_x.TcPOU
(*~
	<docu>
		<summary>
			Encodes the control data into the 256-byte output image (00h command, 06h program, 08h/09h special cycle, 20h parameter request).
		</summary>
	</docu>
~*)
FUNCTION TcoAteqG6_EncodeControl_v_3_5_x : BOOL
VAR_IN_OUT
	inoControl : TcoAteqG6_Control_v_3_5_x;
	inoImage : ARRAY[0..255] OF BYTE;
END_VAR
VAR
	i : INT;
END_VAR

// the whole output image is rewritten every cycle
FOR i := 0 TO 255 DO
	inoImage[i] := 0;
END_FOR
TcoAteqG6_DecodeCommandBits_v_3_5_x(inValue := inoControl.Command, inoBits := inoControl.CommandBits);
TcoAteqG6_SetWord_v_3_5_x(inOffset := 16#00, inValue := inoControl.Command, inoImage := inoImage);
// program number: 1-based in the component, 0-based on the bus
IF inoControl.ProgramNumber >= 1 THEN
	TcoAteqG6_SetWord_v_3_5_x(inOffset := 16#06, inValue := INT_TO_WORD(inoControl.ProgramNumber - 1), inoImage := inoImage);
END_IF
inoImage[16#08] := TcoAteqG6_SpecialCycleToByte_v_3_5_x(inoControl.SpecialCycle);
inoImage[16#09] := inoControl.SpecialCycleInstruction;
// 20h: parameter request - count, then 35 identifiers (22h..67h)
TcoAteqG6_SetWord_v_3_5_x(inOffset := 16#20, inValue := INT_TO_WORD(inoControl.ParameterRequest.Count), inoImage := inoImage);
FOR i := 0 TO 34 DO
	TcoAteqG6_SetWord_v_3_5_x(inOffset := 16#22 + 2 * i, inValue := UINT_TO_WORD(inoControl.ParameterRequest.Ids[i]), inoImage := inoImage);
END_FOR
TcoAteqG6_EncodeControl_v_3_5_x := TRUE;

END_FUNCTION

// ---- POUs/Functions/G6/TcoAteqG6_SetWord_v_3_5_x.TcPOU
(*~
	<docu>
		<summary>
			Writes a little-endian WORD at inOffset.
		</summary>
	</docu>
~*)
FUNCTION TcoAteqG6_SetWord_v_3_5_x : BOOL
VAR_INPUT
	inOffset : INT;
	inValue : WORD;
END_VAR
VAR_IN_OUT
	inoImage : ARRAY[0..255] OF BYTE;
END_VAR

inoImage[inOffset] := WORD_TO_BYTE(inValue AND 16#00FF);
inoImage[inOffset + 1] := WORD_TO_BYTE(SHR(inValue, 8));
TcoAteqG6_SetWord_v_3_5_x := TRUE;

END_FUNCTION

// ---- POUs/Functions/G6/TcoAteqG6_SpecialCycleToByte_v_3_5_x.TcPOU
(*~
	<docu>
		<summary>
			Special cycle to its id byte (output 08h).
		</summary>
	</docu>
~*)
FUNCTION TcoAteqG6_SpecialCycleToByte_v_3_5_x : BYTE
VAR_INPUT
	inValue : eTcoAteqG6_SpecialCycle_v_3_5_x;
END_VAR

CASE inValue OF
	eTcoAteqG6_SpecialCycle_v_3_5_x.AtrLearning: TcoAteqG6_SpecialCycleToByte_v_3_5_x := 1;
	eTcoAteqG6_SpecialCycle_v_3_5_x.CustomUnitLearn: TcoAteqG6_SpecialCycleToByte_v_3_5_x := 4;
	eTcoAteqG6_SpecialCycle_v_3_5_x.CustomUnitCheck: TcoAteqG6_SpecialCycleToByte_v_3_5_x := 5;
	eTcoAteqG6_SpecialCycle_v_3_5_x.PiezoAutoZero: TcoAteqG6_SpecialCycleToByte_v_3_5_x := 9;
	eTcoAteqG6_SpecialCycle_v_3_5_x.RegulatorAdjust: TcoAteqG6_SpecialCycleToByte_v_3_5_x := 13;
	eTcoAteqG6_SpecialCycle_v_3_5_x.CapillaryTemperatureCheck: TcoAteqG6_SpecialCycleToByte_v_3_5_x := 25;
	eTcoAteqG6_SpecialCycle_v_3_5_x.TemperatureCheck: TcoAteqG6_SpecialCycleToByte_v_3_5_x := 26;
	eTcoAteqG6_SpecialCycle_v_3_5_x.AtmPressureCheck: TcoAteqG6_SpecialCycleToByte_v_3_5_x := 27;
	eTcoAteqG6_SpecialCycle_v_3_5_x.P1SensorCheck: TcoAteqG6_SpecialCycleToByte_v_3_5_x := 28;
	eTcoAteqG6_SpecialCycle_v_3_5_x.Flow1Check: TcoAteqG6_SpecialCycleToByte_v_3_5_x := 29;
	eTcoAteqG6_SpecialCycle_v_3_5_x.Flow2Check: TcoAteqG6_SpecialCycleToByte_v_3_5_x := 30;
	eTcoAteqG6_SpecialCycle_v_3_5_x.LinePressureSensorCheck: TcoAteqG6_SpecialCycleToByte_v_3_5_x := 31;
ELSE
	TcoAteqG6_SpecialCycleToByte_v_3_5_x := 0;
END_CASE

END_FUNCTION

// ---- POUs/Functions/G6/TcoAteqG6_IsParameterRequestValid_v_3_5_x.TcPOU
(*~
	<docu>
		<summary>
			TRUE when the request holds 1..35 identifiers.
		</summary>
	</docu>
~*)
FUNCTION TcoAteqG6_IsParameterRequestValid_v_3_5_x : BOOL
VAR_IN_OUT
	inoRequest : TcoAteqG6_ParameterRequest_v_3_5_x;
END_VAR

TcoAteqG6_IsParameterRequestValid_v_3_5_x := inoRequest.Count >= 1 AND inoRequest.Count <= 35;

END_FUNCTION

// ---- POUs/Functions/G6/TcoAteqG6_MapPresetParameters_v_3_5_x.TcPOU
(*~
	<docu>
		<summary>
			Maps a list read with the preset request onto the typed parameter set.
		</summary>
	</docu>
~*)
FUNCTION TcoAteqG6_MapPresetParameters_v_3_5_x : BOOL
VAR_IN_OUT
	inoList : TcoAteqG6_ParameterList_v_3_5_x;
	inoSet : TcoAteqG6_ParameterSet_v_3_5_x;
END_VAR

inoSet.FillTime := TcoAteqG6_ToEngineering_v_3_5_x(TcoAteqG6_TryGetParameterRaw_v_3_5_x(inId := TO_UINT(eTcoAteqG6_ParameterId_v_3_5_x.FillTime), inoList := inoList));
inoSet.StabTime := TcoAteqG6_ToEngineering_v_3_5_x(TcoAteqG6_TryGetParameterRaw_v_3_5_x(inId := TO_UINT(eTcoAteqG6_ParameterId_v_3_5_x.StabTime), inoList := inoList));
inoSet.TestTime := TcoAteqG6_ToEngineering_v_3_5_x(TcoAteqG6_TryGetParameterRaw_v_3_5_x(inId := TO_UINT(eTcoAteqG6_ParameterId_v_3_5_x.TestTime), inoList := inoList));
inoSet.DumpTime := TcoAteqG6_ToEngineering_v_3_5_x(TcoAteqG6_TryGetParameterRaw_v_3_5_x(inId := TO_UINT(eTcoAteqG6_ParameterId_v_3_5_x.DumpTime), inoList := inoList));
inoSet.TestType := TcoAteqG6_ToTestType_v_3_5_x(TcoAteqG6_TryGetParameterRaw_v_3_5_x(inId := TO_UINT(eTcoAteqG6_ParameterId_v_3_5_x.TestType), inoList := inoList));
inoSet.MinFill := TcoAteqG6_ToEngineering_v_3_5_x(TcoAteqG6_TryGetParameterRaw_v_3_5_x(inId := TO_UINT(eTcoAteqG6_ParameterId_v_3_5_x.MinFill), inoList := inoList));
inoSet.MaxFill := TcoAteqG6_ToEngineering_v_3_5_x(TcoAteqG6_TryGetParameterRaw_v_3_5_x(inId := TO_UINT(eTcoAteqG6_ParameterId_v_3_5_x.MaxFill), inoList := inoList));
inoSet.PressureUnit := TcoAteqG6_ToUnit_v_3_5_x(TcoAteqG6_TryGetParameterRaw_v_3_5_x(inId := TO_UINT(eTcoAteqG6_ParameterId_v_3_5_x.PressureUnit), inoList := inoList));
inoSet.TestFail := TcoAteqG6_ToEngineering_v_3_5_x(TcoAteqG6_TryGetParameterRaw_v_3_5_x(inId := TO_UINT(eTcoAteqG6_ParameterId_v_3_5_x.TestFail), inoList := inoList));
inoSet.RefFail := TcoAteqG6_ToEngineering_v_3_5_x(TcoAteqG6_TryGetParameterRaw_v_3_5_x(inId := TO_UINT(eTcoAteqG6_ParameterId_v_3_5_x.RefFail), inoList := inoList));
inoSet.SetFill := TcoAteqG6_ToEngineering_v_3_5_x(TcoAteqG6_TryGetParameterRaw_v_3_5_x(inId := TO_UINT(eTcoAteqG6_ParameterId_v_3_5_x.SetFill), inoList := inoList));
TcoAteqG6_MapPresetParameters_v_3_5_x := TRUE;

END_FUNCTION

// ---- POUs/Functions/G6/TcoAteqG6_TryGetParameterRaw_v_3_5_x.TcPOU
(*~
	<docu>
		<summary>
			Raw value of parameter inId; outFound is FALSE when it is not in the list.
		</summary>
	</docu>
~*)
FUNCTION TcoAteqG6_TryGetParameterRaw_v_3_5_x : DINT
VAR_INPUT
	inId : UINT;
END_VAR
VAR_IN_OUT
	inoList : TcoAteqG6_ParameterList_v_3_5_x;
END_VAR
VAR_OUTPUT
	outFound : BOOL;
END_VAR
VAR
	i : INT;
END_VAR

outFound := FALSE;
FOR i := 0 TO inoList.Count - 1 DO
	IF inoList.Items[i].Id = inId THEN
		TcoAteqG6_TryGetParameterRaw_v_3_5_x := inoList.Items[i].Raw;
		outFound := TRUE;
		RETURN;
	END_IF
END_FOR

END_FUNCTION

// ---- POUs/Functions/G6/TcoAteqG6_ToTestType_v_3_5_x.TcPOU
(*~
	<docu>
		<summary>
			Test type parameter value (code x1000) to test type.
		</summary>
	</docu>
~*)
FUNCTION TcoAteqG6_ToTestType_v_3_5_x : eTcoAteqG6_TestType_v_3_5_x
VAR_INPUT
	inRaw : DINT;
END_VAR

CASE inRaw OF
	0: TcoAteqG6_ToTestType_v_3_5_x := eTcoAteqG6_TestType_v_3_5_x.Invalid;
	1000: TcoAteqG6_ToTestType_v_3_5_x := eTcoAteqG6_TestType_v_3_5_x.Direct;
	2000: TcoAteqG6_ToTestType_v_3_5_x := eTcoAteqG6_TestType_v_3_5_x.Operator;
ELSE
	TcoAteqG6_ToTestType_v_3_5_x := eTcoAteqG6_TestType_v_3_5_x.Unknown;
END_CASE

END_FUNCTION

// ---- POUs/Functions/G6/TcoAteqG6_QueryParameter_v_3_5_x.TcPOU
(*~
	<docu>
		<summary>
			Looks inParameter up in a list that was read.
		</summary>
	</docu>
~*)
FUNCTION TcoAteqG6_QueryParameter_v_3_5_x : BOOL
VAR_INPUT
	inParameter : eTcoAteqG6_ParameterId_v_3_5_x;
END_VAR
VAR_IN_OUT
	inoList : TcoAteqG6_ParameterList_v_3_5_x;
	inoQuery : TcoAteqG6_ParameterQuery_v_3_5_x;
END_VAR

inoQuery.Parameter := inParameter;
inoQuery.Found := FALSE;
inoQuery.Raw := 0;
inoQuery.Value := 0.0;
TcoAteqG6_QueryParameter_v_3_5_x := TRUE;
IF inParameter = eTcoAteqG6_ParameterId_v_3_5_x.None THEN
	RETURN;
END_IF
inoQuery.Raw := TcoAteqG6_TryGetParameterRaw_v_3_5_x(inId := TO_UINT(inParameter), inoList := inoList, outFound => inoQuery.Found);
inoQuery.Value := TcoAteqG6_ToEngineering_v_3_5_x(inoQuery.Raw);

END_FUNCTION

// ---- POUs/Functions/G6/TcoAteqG6_SetDint_v_3_5_x.TcPOU
(*~
	<docu>
		<summary>
			Writes a little-endian LONG at inOffset.
		</summary>
	</docu>
~*)
FUNCTION TcoAteqG6_SetDint_v_3_5_x : BOOL
VAR_INPUT
	inOffset : INT;
	inValue : DINT;
END_VAR
VAR_IN_OUT
	inoImage : ARRAY[0..255] OF BYTE;
END_VAR
VAR
	raw : DWORD;
END_VAR

raw := DINT_TO_DWORD(inValue);
inoImage[inOffset] := DWORD_TO_BYTE(raw);
inoImage[inOffset + 1] := DWORD_TO_BYTE(SHR(raw, 8));
inoImage[inOffset + 2] := DWORD_TO_BYTE(SHR(raw, 16));
inoImage[inOffset + 3] := DWORD_TO_BYTE(SHR(raw, 24));
TcoAteqG6_SetDint_v_3_5_x := TRUE;

END_FUNCTION

// ---- POUs/Prototypes/G6/TcoAteqG6Pn_v_3_5_x.TcPOU
(*~
	<docu>
		<summary>
			ATEQ G6 leak tester (G6 Series - Profinet, fieldbus software 3.5, fieldbus mode 5 "Standard"), PN.
			The interface uses 4 input modules of 64 bytes (slots 1-4) and 4 output modules of 64 bytes (slots 5-8);
			they are mapped to one 256-byte input image and one 256-byte output image. All data are little-endian,
			measured values and parameters are LONG x1000, program numbers are 0-based on the bus and 1-based here.
			Commands use the ATEQ handshake (command bit -> echo -> error word -> release), see TcoAteqG6Task_v_3_5_x.
			Ported from AXOpen AxoG6 v_3_5_x; the hardware-ID bootstrap and the numeric error codes are not ported.
		</summary>
	</docu>
~*)
FUNCTION_BLOCK TcoAteqG6Pn_v_3_5_x EXTENDS TcoIo.TcoPnIoComponent
VAR_INPUT
	inEnable : BOOL;
END_VAR
VAR_IN_OUT
	inoData : TcoAteqG6Pn_IO_v_3_5_x;
END_VAR
VAR
	{attribute addProperty Name "<#Status#>"}
	{attribute clr [ReadOnly()]}
	_status : TcoAteqG6_Status_v_3_5_x;
	{attribute addProperty Name "<#Control#>"}
	_control : TcoAteqG6_Control_v_3_5_x;
	{attribute addProperty Name "<#Config#>"}
	_config : TcoAteqG6_Config_v_3_5_x;
	{attribute addProperty Name "<#PN Error#>"}
	{attribute clr [ReadOnly()]}
	_busError : BOOL;
END_VAR
VAR
	{attribute addProperty Name "<#Reset#>"}
	_resetTask : TcoAteqG6_ResetTask_v_3_5_x(THIS^);

	{attribute addProperty Name "<#Select program#>"}
	_selectProgramTask : TcoAteqG6_SelectProgramTask_v_3_5_x(THIS^);

	{attribute addProperty Name "<#Start test cycle#>"}
	_startCycleTask : TcoAteqG6_StartCycleTask_v_3_5_x(THIS^);

	{attribute addProperty Name "<#Read last result#>"}
	_readLastResultTask : TcoAteqG6_ReadLastResultTask_v_3_5_x(THIS^);

	{attribute addProperty Name "<#Start special cycle#>"}
	_specialCycleTask : TcoAteqG6_SpecialCycleTask_v_3_5_x(THIS^);

	{attribute addProperty Name "<#Read parameters#>"}
	_readParametersTask : TcoAteqG6_ReadParametersTask_v_3_5_x(THIS^);

	{attribute addProperty Name "<#Restore#>"}
	_restoreTask : TcoCore.TcoTask(THIS^);
END_VAR
VAR
	{attribute 'hide'}
	_inputImage : ARRAY[0..255] OF BYTE;
	{attribute 'hide'}
	_outputImage : ARRAY[0..255] OF BYTE;
	{attribute 'hide'}
	_sb : TcoCore.StringBuilder;
END_VAR

IF NOT __ISVALIDREF(inoData) THEN
	Messenger.Post('Invalid reference', TcoCore.eMessageCategory.ProgrammingError);
	RETURN;
END_IF

SUPER^(inPnIoBoxState := THIS^.inoData.PnIoBoxState, inPnIoBoxDiag := THIS^.inoData.PnIoBoxDiag);
_busError := NOT _profinetReady;

UpdateStatus();

// Reset is never blocked and aborts any other running command
_resetTask.Enabled := TRUE;
IF _resetTask.Busy THEN
	AbortCommandTasks();
END_IF
_resetTask(inoConfig := _config, inoControl := _control, inoStatus := _status, inoImage := _inputImage);

// one command at a time: every other command is disabled while any command task is busy
_selectProgramTask.Enabled := NOT (_resetTask.Busy OR _startCycleTask.Busy OR _readLastResultTask.Busy OR _specialCycleTask.Busy OR _readParametersTask.Busy);
_selectProgramTask(inoConfig := _config, inoControl := _control, inoStatus := _status, inoImage := _inputImage);

_startCycleTask.Enabled := NOT (_resetTask.Busy OR _selectProgramTask.Busy OR _readLastResultTask.Busy OR _specialCycleTask.Busy OR _readParametersTask.Busy);
_startCycleTask(inoConfig := _config, inoControl := _control, inoStatus := _status, inoImage := _inputImage);

_readLastResultTask.Enabled := NOT (_resetTask.Busy OR _selectProgramTask.Busy OR _startCycleTask.Busy OR _specialCycleTask.Busy OR _readParametersTask.Busy);
_readLastResultTask(inoConfig := _config, inoControl := _control, inoStatus := _status, inoImage := _inputImage);

_specialCycleTask.Enabled := NOT (_resetTask.Busy OR _selectProgramTask.Busy OR _startCycleTask.Busy OR _readLastResultTask.Busy OR _readParametersTask.Busy);
_specialCycleTask(inoConfig := _config, inoControl := _control, inoStatus := _status, inoImage := _inputImage);

_readParametersTask.Enabled := NOT (_resetTask.Busy OR _selectProgramTask.Busy OR _startCycleTask.Busy OR _readLastResultTask.Busy OR _specialCycleTask.Busy);
_readParametersTask(inoConfig := _config, inoControl := _control, inoStatus := _status, inoImage := _inputImage);

//*************RESTORE********************
_restoreTask.Enabled := TRUE;
IF _restoreTask.Execute() THEN
	Restore();
	_restoreTask.DoneWhen(TRUE);
END_IF
//****************************************

UpdateControl();

(*~
	<docu>
		<summary>
			Gets the configuration of the instrument.
		</summary>
	</docu>
~*)
PROPERTY Config : REFERENCE TO TcoAteqG6_Config_v_3_5_x
GET
Config REF= _config;
END_GET
END_PROPERTY

PROPERTY PUBLIC Control : REFERENCE TO TcoAteqG6_Control_v_3_5_x
GET
Control REF= _control;
END_GET
END_PROPERTY

(*~
	<docu>
		<summary>
			Gets the status of the instrument (live state, last result, parameters).
		</summary>
	</docu>
~*)
PROPERTY Status : REFERENCE TO TcoAteqG6_Status_v_3_5_x
GET
Status REF= _status;
END_GET
END_PROPERTY

METHOD FB_init : BOOL
VAR_INPUT
	bInitRetains : BOOL; // if TRUE, the retain variables are initialized (warm start / cold start)
	bInCopyCode : BOOL;  // if TRUE, the instance afterwards gets moved into the copy code (online change)
	ParentObject : ITcoObject;
END_VAR
END_METHOD

METHOD INTERNAL AbortCommandTasks
_selectProgramTask.Abort();
_startCycleTask.Abort();
_readLastResultTask.Abort();
_specialCycleTask.Abort();
_readParametersTask.Abort();
END_METHOD

METHOD INTERNAL CommandTaskBusy : BOOL
CommandTaskBusy := _resetTask.Busy OR _selectProgramTask.Busy OR _startCycleTask.Busy OR _readLastResultTask.Busy OR _specialCycleTask.Busy OR _readParametersTask.Busy;
END_METHOD

(*~
	<docu>
		<summary>
			Restores this instance to the Ready state. Can be called explicitly or from within one of the restore mechanisms.
		</summary>
	</docu>
~*)
METHOD Restore : ITcoRestorable
RestoreTasks();
_control.Command := 0;
_status.LastCommandError := 0;
_status.ActionDescription := '<#Restore has been executed.#>';
END_METHOD

METHOD INTERNAL RestoreTasks
_resetTask.Restore();
_selectProgramTask.Restore();
_startCycleTask.Restore();
_readLastResultTask.Restore();
_specialCycleTask.Restore();
_readParametersTask.Restore();
END_METHOD

(*~
	<docu>
		<summary>
			Custom service (manual, maintenance) logic.
		</summary>
	</docu>
~*)
METHOD PROTECTED ServiceMode
END_METHOD

(*~
	<docu>
		<summary>
			Copies the 4 input modules into the 256-byte input image and decodes the live state.
		</summary>
	</docu>
~*)
METHOD INTERNAL UpdateStatus
MEMCPY(destAddr := ADR(_inputImage[0]), srcAddr := ADR(inoData.In.In1), n := 64);
MEMCPY(destAddr := ADR(_inputImage[64]), srcAddr := ADR(inoData.In.In2), n := 64);
MEMCPY(destAddr := ADR(_inputImage[128]), srcAddr := ADR(inoData.In.In3), n := 64);
MEMCPY(destAddr := ADR(_inputImage[192]), srcAddr := ADR(inoData.In.In4), n := 64);

TcoAteqG6_DecodeState_v_3_5_x(inoImage := _inputImage, inoState := _status.State);
_status.Ready := _status.State.StatusBits.CycleEnd AND NOT _status.State.CommandRunning;
_status.LastPass := _status.LastResult.Valid AND _status.LastResult.Pass;
END_METHOD

(*~
	<docu>
		<summary>
			Encodes the control data into the 256-byte output image and copies it to the 4 output modules.
		</summary>
	</docu>
~*)
METHOD INTERNAL UpdateControl
TcoAteqG6_EncodeControl_v_3_5_x(inoControl := _control, inoImage := _outputImage);

MEMCPY(destAddr := ADR(inoData.Out.Out1), srcAddr := ADR(_outputImage[0]), n := 64);
MEMCPY(destAddr := ADR(inoData.Out.Out2), srcAddr := ADR(_outputImage[64]), n := 64);
MEMCPY(destAddr := ADR(inoData.Out.Out3), srcAddr := ADR(_outputImage[128]), n := 64);
MEMCPY(destAddr := ADR(inoData.Out.Out4), srcAddr := ADR(_outputImage[192]), n := 64);
END_METHOD

(*~
	<docu>
		<summary>
			Resets the instrument. Aborts any other running command.
		</summary>
	</docu>
~*)
METHOD PUBLIC Reset : TcoCore.ITcoTaskStatus
AbortCommandTasks();
Reset := _resetTask.Invoke();
END_METHOD

(*~
	<docu>
		<summary>
			Selects program inProgram (1-128, as shown on the instrument display).
		</summary>
	</docu>
~*)
METHOD PUBLIC SelectProgram : TcoCore.ITcoTaskStatus
VAR_INPUT
	inProgram : INT;
END_VAR
IF _selectProgramTask.Busy OR NOT CommandTaskBusy() THEN
	_control.ProgramNumber := inProgram;
END_IF
SelectProgram := _selectProgramTask.Invoke();
END_METHOD

(*~
	<docu>
		<summary>
			Runs a complete test cycle on program inProgram (1-128) and reads its result into Status.LastResult.
		</summary>
	</docu>
~*)
METHOD PUBLIC StartCycle : TcoCore.ITcoTaskStatus
VAR_INPUT
	inProgram : INT;
END_VAR
IF _startCycleTask.Busy OR NOT CommandTaskBusy() THEN
	_control.ProgramNumber := inProgram;
END_IF
StartCycle := _startCycleTask.Invoke();
END_METHOD

METHOD PUBLIC ReadLastResult : TcoCore.ITcoTaskStatus
ReadLastResult := _readLastResultTask.Invoke();
END_METHOD

(*~
	<docu>
		<summary>
			Runs special cycle inSpecialCycle with instruction inInstruction on the currently selected program.
		</summary>
	</docu>
~*)
METHOD PUBLIC SpecialCycle : TcoCore.ITcoTaskStatus
VAR_INPUT
	inSpecialCycle : eTcoAteqG6_SpecialCycle_v_3_5_x;
	inInstruction : BYTE;
END_VAR
IF _specialCycleTask.Busy OR NOT CommandTaskBusy() THEN
	_control.SpecialCycle := inSpecialCycle;
	_control.SpecialCycleInstruction := inInstruction;
END_IF
SpecialCycle := _specialCycleTask.Invoke();
END_METHOD

(*~
	<docu>
		<summary>
			Reads the parameters listed in inoRequest (1-35 identifiers) into Status.Parameters.
		</summary>
	</docu>
~*)
METHOD PUBLIC ReadParameters : TcoCore.ITcoTaskStatus
VAR_IN_OUT
	inoRequest : TcoAteqG6_ParameterRequest_v_3_5_x;
END_VAR
IF _readParametersTask.Busy OR NOT CommandTaskBusy() THEN
	_control.ParameterRequest := inoRequest;
END_IF
ReadParameters := _readParametersTask.InvokeWithParams(inMapToPreset := FALSE);
END_METHOD

(*~
	<docu>
		<summary>
			Reads the preset parameters (times, test type, fill levels, reject levels) into Status.ParameterSet.
		</summary>
	</docu>
~*)
METHOD PUBLIC ReadPresetParameters : TcoCore.ITcoTaskStatus
IF _readParametersTask.Busy OR NOT CommandTaskBusy() THEN
	TcoAteqG6_BuildPresetRequest_v_3_5_x(inoRequest := _control.ParameterRequest);
END_IF
ReadPresetParameters := _readParametersTask.InvokeWithParams(inMapToPreset := TRUE);
END_METHOD

(*~
	<docu>
		<summary>
			Reads one parameter; the value is in Status.ParameterQuery.
		</summary>
	</docu>
~*)
METHOD PUBLIC ReadParameter : TcoCore.ITcoTaskStatus
VAR_INPUT
	inParameter : eTcoAteqG6_ParameterId_v_3_5_x;
END_VAR
IF _readParametersTask.Busy OR NOT CommandTaskBusy() THEN
	TcoAteqG6_ClearParameterRequest_v_3_5_x(inoRequest := _control.ParameterRequest);
	TcoAteqG6_AddParameterToRequest_v_3_5_x(inParameter := inParameter, inoRequest := _control.ParameterRequest);
	_control.QueryParameter := inParameter;
END_IF
ReadParameter := _readParametersTask.InvokeWithParams(inMapToPreset := FALSE);
END_METHOD

PROPERTY ResetTask : TcoCore.ITcoTaskStatus
GET
ResetTask := _resetTask;
END_GET
END_PROPERTY

PROPERTY SelectProgramTask : TcoCore.ITcoTaskStatus
GET
SelectProgramTask := _selectProgramTask;
END_GET
END_PROPERTY

PROPERTY StartCycleTask : TcoCore.ITcoTaskStatus
GET
StartCycleTask := _startCycleTask;
END_GET
END_PROPERTY

PROPERTY ReadLastResultTask : TcoCore.ITcoTaskStatus
GET
ReadLastResultTask := _readLastResultTask;
END_GET
END_PROPERTY

PROPERTY SpecialCycleTask : TcoCore.ITcoTaskStatus
GET
SpecialCycleTask := _specialCycleTask;
END_GET
END_PROPERTY

PROPERTY ReadParametersTask : TcoCore.ITcoTaskStatus
GET
ReadParametersTask := _readParametersTask;
END_GET
END_PROPERTY

END_FUNCTION_BLOCK

// ---- POUs/Prototypes/MeasurementTasks/G6_v_3_5_x/TcoAteqG6_ResetTask_v_3_5_x.TcPOU
(*~
	<docu>
		<summary>
			Reset command (command bit 0). Never blocked; aborts any other running command.
		</summary>
	</docu>
~*)
FUNCTION_BLOCK TcoAteqG6_ResetTask_v_3_5_x EXTENDS TcoAteqG6Task_v_3_5_x

IF Execute() THEN
	IF CheckReferences() THEN
		// AX step 0: reset handshake
		IF _progress = 0 THEN
			inoStatus.ActionDescription := '<#Resetting instrument#>';
			IF Handshake(MASK_RESET) THEN
				GoTo(100);
			END_IF
		END_IF

		// AX step 100
		IF _progress = 100 THEN
			inoStatus.ActionDescription := '<#Instrument reset#>';
			DoneWhen(TRUE);
		END_IF
		Supervise();
	END_IF
END_IF

IF THIS^.Error AND NOT _errorMessage.Pinned THEN
	THIS^.Restore();
END_IF

METHOD FB_init : BOOL
VAR_INPUT
	bInitRetains : BOOL; // if TRUE, the retain variables are initialized (warm start / cold start)
	bInCopyCode : BOOL;  // if TRUE, the instance afterwards gets moved into the copy code (online change)
	ParentObject : ITcoObject;
END_VAR
END_METHOD

END_FUNCTION_BLOCK

// ---- POUs/Prototypes/MeasurementTasks/G6_v_3_5_x/TcoAteqG6Task_v_3_5_x.TcPOU
(*~
	<docu>
		<summary>
			Base of every ATEQ G6 command task. Owns the command handshake (manual p. 56):
			own echo low -> raise the command bit (single rising edge) -> acknowledged (error word FFFFh or echo set) ->
			completed (error word <> FFFFh; 0 = ok, otherwise failed) -> drop the command bit -> echo low.
			Every wait is bounded by Config.CommandTimeout. The command bit is always dropped on done, error, abort and
			restore - the instrument only reacts to rising edges, so a bit left high would make it miss the next command.
		</summary>
	</docu>
~*)
FUNCTION_BLOCK PUBLIC ABSTRACT TcoAteqG6Task_v_3_5_x EXTENDS TcoCore.TcoTask
VAR_IN_OUT
	inoConfig : TcoAteqG6_Config_v_3_5_x;
	inoControl : TcoAteqG6_Control_v_3_5_x;
	inoStatus : TcoAteqG6_Status_v_3_5_x;
	inoImage : ARRAY[0..255] OF BYTE;
END_VAR
VAR
	_errorMessage : TcoCore.TcoMessenger(THIS^);
	{attribute 'hide'}
	_progress : INT := 0;
	{attribute 'hide'}
	_hsStep : INT := 0;
	{attribute 'hide'}
	_activeMask : WORD;
	{attribute 'hide'}
	_cycleRunningSeen : BOOL;
	{attribute 'hide'}
	_failText : STRING(254);
	{attribute 'hide'}
	_stepTimer : TON;
	{attribute 'hide'}
	_hsTimer : TON;
	{attribute 'hide'}
	_infoTimer : TON;
	{attribute 'hide'}
	_errorTimer : TON;
	{attribute 'hide'}
	_varInfo : __SYSTEM.VAR_INFO;
	{attribute 'hide'}
	_sb : TcoCore.StringBuilder;
END_VAR
VAR CONSTANT
	MASK_RESET : WORD := 16#0001;
	MASK_START : WORD := 16#0002;
	MASK_SPECIAL_CYCLE : WORD := 16#0006; // Start + Special cycle, sent together
	MASK_PROGRAM_SELECTION : WORD := 16#0008;
	MASK_READ_PARAMETERS : WORD := 16#0020;
	MASK_READ_LAST_RESULT : WORD := 16#8000;
END_VAR

METHOD CallTimers
VAR_INPUT
	inValue : BOOL;
END_VAR
IF __ISVALIDREF(inoConfig) AND THIS^.inoConfig.ErrorTime <> T#0S OR NOT inValue THEN
	_errorTimer(IN := inValue, PT := THIS^.inoConfig.ErrorTime);
END_IF
IF __ISVALIDREF(inoConfig) AND THIS^.inoConfig.InfoTime <> T#0S OR NOT inValue THEN
	_infoTimer(IN := inValue, PT := THIS^.inoConfig.InfoTime);
END_IF
END_METHOD

(*~
	<docu>
		<summary>
			Checks the references to the config, control, status and input image. Returns TRUE when all of them are valid.
		</summary>
	</docu>
~*)
METHOD PROTECTED CheckReferences : BOOL
IF NOT __ISVALIDREF(inoControl) THEN
	_varInfo := __VARINFO(inoControl);
	Messenger.Programming(_sb.Clear().Append('<#Invalid reference: #>').Append(_varInfo.Symbol).ToString()).Pin();
ELSIF NOT __ISVALIDREF(inoConfig) THEN
	_varInfo := __VARINFO(inoConfig);
	Messenger.Programming(_sb.Clear().Append('<#Invalid reference: #>').Append(_varInfo.Symbol).ToString()).Pin();
ELSIF NOT __ISVALIDREF(inoStatus) THEN
	_varInfo := __VARINFO(inoStatus);
	Messenger.Programming(_sb.Clear().Append('<#Invalid reference: #>').Append(_varInfo.Symbol).ToString()).Pin();
ELSIF NOT __ISVALIDREF(inoImage) THEN
	_varInfo := __VARINFO(inoImage);
	Messenger.Programming(_sb.Clear().Append('<#Invalid reference: #>').Append(_varInfo.Symbol).ToString()).Pin();
ELSE
	CheckReferences := TRUE;
END_IF
END_METHOD

METHOD PROTECTED CommandTimeout : TIME
IF __ISVALIDREF(inoConfig) AND THIS^.inoConfig.CommandTimeout > T#0S THEN
	CommandTimeout := THIS^.inoConfig.CommandTimeout;
ELSE
	CommandTimeout := T#5S;
END_IF
END_METHOD

METHOD PROTECTED CycleTimeout : TIME
IF __ISVALIDREF(inoConfig) AND THIS^.inoConfig.CycleTimeout > T#0S THEN
	CycleTimeout := THIS^.inoConfig.CycleTimeout;
ELSE
	CycleTimeout := T#60S;
END_IF
END_METHOD

(*~
	<docu>
		<summary>
			Puts the task into error with the text inText, keeps the command error word and drops the command bit.
		</summary>
	</docu>
~*)
METHOD PROTECTED Fail
VAR_INPUT
	inText : STRING(254);
END_VAR
_failText := inText;
IF __ISVALIDREF(inoStatus) THEN
	THIS^.inoStatus.LastCommandError := THIS^.inoStatus.State.Error.Raw;
END_IF
ReleaseCommand();
_hsStep := 0;
THIS^.ThrowWhen(TRUE);
END_METHOD

(*~
	<docu>
		<summary>
			Moves to inStep and restarts the step timer.
		</summary>
	</docu>
~*)
METHOD PROTECTED GoTo
VAR_INPUT
	inStep : INT;
END_VAR
_stepTimer(IN := FALSE);
_progress := inStep;
END_METHOD

(*~
	<docu>
		<summary>
			Runs one command handshake for inMask. Returns TRUE in the cycle the handshake finished successfully;
			on any failure the task is put into error.
		</summary>
	</docu>
~*)
METHOD PROTECTED Handshake : BOOL
VAR_INPUT
	inMask : WORD;
END_VAR
// 0: the instrument must not still echo this command (previous one not released)
IF _hsStep = 0 THEN
	_hsTimer(IN := TRUE, PT := CommandTimeout());
	IF (inoStatus.State.Echo.Raw AND inMask) = 0 THEN
		_hsTimer(IN := FALSE);
		_hsStep := 1;
	ELSIF _hsTimer.Q THEN
		Fail('<#Instrument still echoes the previous command. Reset the instrument, then restore the component.#>');
		RETURN;
	END_IF
END_IF

// 1: raise the command bit - a single rising edge
IF _hsStep = 1 THEN
	_activeMask := inMask;
	inoControl.Command := inoControl.Command OR inMask;
	_hsStep := 2;
END_IF

// 2: acknowledged - command running (FFFFh) or already echoed
IF _hsStep = 2 THEN
	_hsTimer(IN := TRUE, PT := CommandTimeout());
	IF inoStatus.State.Error.Raw = 16#FFFF OR (inoStatus.State.Echo.Raw AND inMask) = inMask THEN
		_hsTimer(IN := FALSE);
		_hsStep := 3;
	ELSIF _hsTimer.Q THEN
		Fail('<#Command was not acknowledged by the instrument. Check the PROFINET connection and fieldbus mode 5 Standard.#>');
		RETURN;
	END_IF
END_IF

// 3: completed - error word left FFFFh; 0 = success, anything else = failed
IF _hsStep = 3 THEN
	_hsTimer(IN := TRUE, PT := CommandTimeout());
	IF inoStatus.State.Error.Raw <> 16#FFFF AND (inoStatus.State.Echo.Raw AND inMask) = inMask THEN
		_hsTimer(IN := FALSE);
		IF inoStatus.State.Error.Raw <> 0 THEN
			Fail('<#Instrument reported a command error. See LastCommandError: the set bit names the failed command.#>');
			RETURN;
		END_IF
		_hsStep := 4;
	ELSIF _hsTimer.Q THEN
		Fail('<#Command was not completed by the instrument. Check the instrument display for a running menu or alarm.#>');
		RETURN;
	END_IF
END_IF

// 4: drop the command bit
IF _hsStep = 4 THEN
	ReleaseCommand();
	_hsStep := 5;
END_IF

// 5: echo released
IF _hsStep = 5 THEN
	_hsTimer(IN := TRUE, PT := CommandTimeout());
	IF (inoStatus.State.Echo.Raw AND inMask) = 0 THEN
		_hsTimer(IN := FALSE);
		_hsStep := 0;
		Handshake := TRUE;
	ELSIF _hsTimer.Q THEN
		Fail('<#Instrument did not release the command echo. Reset the instrument, then restore the component.#>');
		RETURN;
	END_IF
END_IF
END_METHOD

(*~
	<docu>
		<summary>
			Waits for a full cycle after a start command: CycleEnd must be seen FALSE (cycle running, within
			Config.CommandTimeout of the start) and then TRUE again (within Config.CycleTimeout). Call it every cycle from
			the moment the start bit is raised, so a cycle that starts during the handshake is not missed.
			Returns TRUE when the cycle ended.
		</summary>
	</docu>
~*)
METHOD PROTECTED ObserveCycle : BOOL
VAR_INPUT
	inWaiting : BOOL; // FALSE while the start handshake is still running
END_VAR
IF NOT inoStatus.State.StatusBits.CycleEnd THEN
	_cycleRunningSeen := TRUE;
END_IF
IF NOT inWaiting THEN
	RETURN;
END_IF
IF NOT _cycleRunningSeen THEN
	IF StepElapsed(CommandTimeout()) THEN
		Fail('<#Test cycle did not start. Check the instrument for alarms and that the program is valid.#>');
	END_IF
ELSIF inoStatus.State.StatusBits.CycleEnd THEN
	ObserveCycle := TRUE;
ELSIF StepElapsed(CycleTimeout()) THEN
	Fail('<#Test cycle did not end within Config.CycleTimeout.#>');
END_IF
END_METHOD

METHOD PROTECTED ReleaseCommand
IF __ISVALIDREF(inoControl) AND _activeMask <> 0 THEN
	THIS^.inoControl.Command := THIS^.inoControl.Command AND NOT _activeMask;
END_IF
_activeMask := 0;
END_METHOD

(*~
	<docu>
		<summary>
			TRUE when the current step has been active longer than inLimit.
		</summary>
	</docu>
~*)
METHOD PROTECTED StepElapsed : BOOL
VAR_INPUT
	inLimit : TIME;
END_VAR
_stepTimer(IN := TRUE, PT := inLimit);
StepElapsed := _stepTimer.Q;
END_METHOD

(*~
	<docu>
		<summary>
			Per-cycle bookkeeping: progress information after Config.InfoTime and the optional task timeout Config.ErrorTime.
		</summary>
	</docu>
~*)
METHOD PROTECTED Supervise
CallTimers(TRUE);
THIS^.Messenger.OnCondition(_infoTimer.Q).Info(inoStatus.ActionDescription);
IF _errorTimer.Q THEN
	Fail('<#Task time exceeded (Config.ErrorTime).#>');
END_IF
END_METHOD

METHOD PROTECTED OnAbort
ReleaseCommand();
_hsStep := 0;
IF __ISVALIDREF(inoStatus) THEN THIS^.inoStatus.ActionDescription := '<#Command was aborted.#>'; END_IF
END_METHOD

METHOD PROTECTED OnDone
ReleaseCommand();
_progress := 0;
END_METHOD

METHOD PROTECTED OnError
ReleaseCommand();
IF __ISVALIDREF(inoStatus) THEN THIS^.inoStatus.ActionDescription := _failText; END_IF
THIS^._errorMessage.Error(_sb.Clear().Append(_failText).Append('<# To restore acknowledge this alarm.#>').ToString()).Pin();
END_METHOD

METHOD PROTECTED OnStart
ReleaseCommand();
_progress := 0;
_hsStep := 0;
_cycleRunningSeen := FALSE;
_failText := '';
_stepTimer(IN := FALSE);
_hsTimer(IN := FALSE);
CallTimers(FALSE);
IF __ISVALIDREF(inoStatus) THEN THIS^.inoStatus.LastCommandError := 0; END_IF
END_METHOD

(*~
	<docu>
		<summary>
			Restores this instance to the Ready state and drops its command bit.
		</summary>
	</docu>
~*)
METHOD Restore : ITcoRestorable
SUPER^.Restore();
ReleaseCommand();
_progress := 0;
_hsStep := 0;
_stepTimer(IN := FALSE);
_hsTimer(IN := FALSE);
CallTimers(FALSE);
Messenger.UnPin();
_errorMessage.UnPin();
END_METHOD

END_FUNCTION_BLOCK

// ---- POUs/Prototypes/MeasurementTasks/G6_v_3_5_x/TcoAteqG6_SelectProgramTask_v_3_5_x.TcPOU
(*~
	<docu>
		<summary>
			Program selection (command bit 3) of Control.ProgramNumber, then checks that the instrument switched to it.
		</summary>
	</docu>
~*)
FUNCTION_BLOCK TcoAteqG6_SelectProgramTask_v_3_5_x EXTENDS TcoAteqG6Task_v_3_5_x

IF Execute() THEN
	IF CheckReferences() THEN
		// AX step 0: valid program number
		IF _progress = 0 THEN
			inoStatus.ActionDescription := '<#Checking program number#>';
			IF inoControl.ProgramNumber < 1 OR inoControl.ProgramNumber > 128 THEN
				Fail('<#Program number out of range (1-128). Pass the program number as shown on the instrument display.#>');
			ELSE
				GoTo(10);
			END_IF
		END_IF

		// AX step 10: select the program
		IF _progress = 10 THEN
			inoStatus.ActionDescription := '<#Selecting program#>';
			IF Handshake(MASK_PROGRAM_SELECTION) THEN
				GoTo(20);
			END_IF
		END_IF

		// AX step 20: the instrument reports the requested program
		IF _progress = 20 THEN
			inoStatus.ActionDescription := '<#Verifying selected program#>';
			IF inoStatus.State.CurrentProgram = inoControl.ProgramNumber THEN
				GoTo(100);
			ELSIF StepElapsed(CommandTimeout()) THEN
				Fail('<#Instrument did not switch to the requested program. Check that the program exists on the instrument.#>');
			END_IF
		END_IF

		// AX step 100
		IF _progress = 100 THEN
			inoStatus.ActionDescription := '<#Program selected#>';
			DoneWhen(TRUE);
		END_IF
		Supervise();
	END_IF
END_IF

IF THIS^.Error AND NOT _errorMessage.Pinned THEN
	THIS^.Restore();
END_IF

METHOD FB_init : BOOL
VAR_INPUT
	bInitRetains : BOOL; // if TRUE, the retain variables are initialized (warm start / cold start)
	bInCopyCode : BOOL;  // if TRUE, the instance afterwards gets moved into the copy code (online change)
	ParentObject : ITcoObject;
END_VAR
END_METHOD

END_FUNCTION_BLOCK

// ---- POUs/Prototypes/MeasurementTasks/G6_v_3_5_x/TcoAteqG6_StartCycleTask_v_3_5_x.TcPOU
(*~
	<docu>
		<summary>
			Complete test cycle on Control.ProgramNumber: select the program, start, wait for the cycle to run and end, then read the last result. A result whose program number differs from the requested one is refused as stale. The results FIFO is never reset.
		</summary>
	</docu>
~*)
FUNCTION_BLOCK TcoAteqG6_StartCycleTask_v_3_5_x EXTENDS TcoAteqG6Task_v_3_5_x

IF Execute() THEN
	IF CheckReferences() THEN
		// AX step 0: preconditions - valid program, instrument at rest (cycle end)
		IF _progress = 0 THEN
			inoStatus.ActionDescription := '<#Waiting for instrument ready#>';
			IF inoControl.ProgramNumber < 1 OR inoControl.ProgramNumber > 128 THEN
				Fail('<#Program number out of range (1-128). Pass the program number as shown on the instrument display.#>');
			ELSIF inoStatus.State.StatusBits.CycleEnd THEN
				GoTo(10);
			ELSIF StepElapsed(CommandTimeout()) THEN
				Fail('<#Instrument is not ready (no cycle end). Wait for the running cycle to finish or reset the instrument.#>');
			END_IF
		END_IF

		// AX step 10: select the program
		IF _progress = 10 THEN
			inoStatus.ActionDescription := '<#Selecting program#>';
			IF Handshake(MASK_PROGRAM_SELECTION) THEN
				GoTo(20);
			END_IF
		END_IF

		// AX step 20: the instrument reports the requested program
		IF _progress = 20 THEN
			inoStatus.ActionDescription := '<#Verifying selected program#>';
			IF inoStatus.State.CurrentProgram = inoControl.ProgramNumber THEN
				_cycleRunningSeen := FALSE;
				GoTo(30);
			ELSIF StepElapsed(CommandTimeout()) THEN
				Fail('<#Instrument did not switch to the requested program. Check that the program exists on the instrument.#>');
			END_IF
		END_IF

		// AX step 30: start; the cycle may already begin while the handshake runs
		IF _progress = 30 THEN
			inoStatus.ActionDescription := '<#Starting test cycle#>';
			ObserveCycle(inWaiting := FALSE);
			IF Handshake(MASK_START) THEN
				GoTo(40);
			END_IF
		END_IF

		// AX step 40: cycle runs (cycle end FALSE) and ends (cycle end TRUE)
		IF _progress = 40 THEN
			inoStatus.ActionDescription := '<#Test cycle running#>';
			IF ObserveCycle(inWaiting := TRUE) THEN
				GoTo(50);
			END_IF
		END_IF

		// AX step 50: read the last result
		IF _progress = 50 THEN
			inoStatus.ActionDescription := '<#Reading last result#>';
			IF Handshake(MASK_READ_LAST_RESULT) THEN
				TcoAteqG6_DecodeLastResult_v_3_5_x(inoImage := inoImage, inoResult := inoStatus.LastResult);
				GoTo(60);
			END_IF
		END_IF

		// AX step 60: the result belongs to this cycle's program
		IF _progress = 60 THEN
			IF inoStatus.LastResult.ProgramNo = inoControl.ProgramNumber THEN
				GoTo(100);
			ELSE
				inoStatus.LastResult.Valid := FALSE;
				Fail('<#Last result does not belong to the requested program. A stale result was read.#>');
			END_IF
		END_IF

		// AX step 100
		IF _progress = 100 THEN
			inoStatus.ActionDescription := '<#Test cycle finished#>';
			DoneWhen(TRUE);
		END_IF
		Supervise();
	END_IF
END_IF

IF THIS^.Error AND NOT _errorMessage.Pinned THEN
	THIS^.Restore();
END_IF

METHOD FB_init : BOOL
VAR_INPUT
	bInitRetains : BOOL; // if TRUE, the retain variables are initialized (warm start / cold start)
	bInCopyCode : BOOL;  // if TRUE, the instance afterwards gets moved into the copy code (online change)
	ParentObject : ITcoObject;
END_VAR
END_METHOD

METHOD PROTECTED OnStart
SUPER^.OnStart();
IF __ISVALIDREF(inoStatus) THEN
	TcoAteqG6_ClearLastResult_v_3_5_x(inoResult := THIS^.inoStatus.LastResult);
END_IF
END_METHOD

END_FUNCTION_BLOCK

// ---- POUs/Prototypes/MeasurementTasks/G6_v_3_5_x/TcoAteqG6_ReadLastResultTask_v_3_5_x.TcPOU
(*~
	<docu>
		<summary>
			Read last result (command bit 15) and decode the exchange zone into Status.LastResult.
		</summary>
	</docu>
~*)
FUNCTION_BLOCK TcoAteqG6_ReadLastResultTask_v_3_5_x EXTENDS TcoAteqG6Task_v_3_5_x

IF Execute() THEN
	IF CheckReferences() THEN
		// AX step 0: read the last result
		IF _progress = 0 THEN
			inoStatus.ActionDescription := '<#Reading last result#>';
			IF Handshake(MASK_READ_LAST_RESULT) THEN
				TcoAteqG6_DecodeLastResult_v_3_5_x(inoImage := inoImage, inoResult := inoStatus.LastResult);
				GoTo(100);
			END_IF
		END_IF

		// AX step 100
		IF _progress = 100 THEN
			inoStatus.ActionDescription := '<#Last result read#>';
			DoneWhen(TRUE);
		END_IF
		Supervise();
	END_IF
END_IF

IF THIS^.Error AND NOT _errorMessage.Pinned THEN
	THIS^.Restore();
END_IF

METHOD FB_init : BOOL
VAR_INPUT
	bInitRetains : BOOL; // if TRUE, the retain variables are initialized (warm start / cold start)
	bInCopyCode : BOOL;  // if TRUE, the instance afterwards gets moved into the copy code (online change)
	ParentObject : ITcoObject;
END_VAR
END_METHOD

METHOD PROTECTED OnStart
SUPER^.OnStart();
IF __ISVALIDREF(inoStatus) THEN
	TcoAteqG6_ClearLastResult_v_3_5_x(inoResult := THIS^.inoStatus.LastResult);
END_IF
END_METHOD

END_FUNCTION_BLOCK

// ---- POUs/Prototypes/MeasurementTasks/G6_v_3_5_x/TcoAteqG6_SpecialCycleTask_v_3_5_x.TcPOU
(*~
	<docu>
		<summary>
			Special cycle Control.SpecialCycle (id at output 08h, instruction at 09h), started with the Start and Special cycle bits together (manual pp. 58-59), then waits for the cycle end. Runs on the currently selected program.
		</summary>
	</docu>
~*)
FUNCTION_BLOCK TcoAteqG6_SpecialCycleTask_v_3_5_x EXTENDS TcoAteqG6Task_v_3_5_x

IF Execute() THEN
	IF CheckReferences() THEN
		// AX step 0: preconditions - special cycle selected, instrument at rest
		IF _progress = 0 THEN
			inoStatus.ActionDescription := '<#Waiting for instrument ready#>';
			IF inoControl.SpecialCycle = eTcoAteqG6_SpecialCycle_v_3_5_x.None THEN
				Fail('<#No special cycle selected.#>');
			ELSIF inoStatus.State.StatusBits.CycleEnd THEN
				_cycleRunningSeen := FALSE;
				GoTo(10);
			ELSIF StepElapsed(CommandTimeout()) THEN
				Fail('<#Instrument is not ready (no cycle end). Wait for the running cycle to finish or reset the instrument.#>');
			END_IF
		END_IF

		// AX step 10: start the special cycle
		IF _progress = 10 THEN
			inoStatus.ActionDescription := '<#Starting special cycle#>';
			ObserveCycle(inWaiting := FALSE);
			IF Handshake(MASK_SPECIAL_CYCLE) THEN
				GoTo(20);
			END_IF
		END_IF

		// AX step 20: cycle runs and ends
		IF _progress = 20 THEN
			inoStatus.ActionDescription := '<#Special cycle running#>';
			IF ObserveCycle(inWaiting := TRUE) THEN
				GoTo(100);
			END_IF
		END_IF

		// AX step 100
		IF _progress = 100 THEN
			inoStatus.ActionDescription := '<#Special cycle finished#>';
			DoneWhen(TRUE);
		END_IF
		Supervise();
	END_IF
END_IF

IF THIS^.Error AND NOT _errorMessage.Pinned THEN
	THIS^.Restore();
END_IF

METHOD FB_init : BOOL
VAR_INPUT
	bInitRetains : BOOL; // if TRUE, the retain variables are initialized (warm start / cold start)
	bInCopyCode : BOOL;  // if TRUE, the instance afterwards gets moved into the copy code (online change)
	ParentObject : ITcoObject;
END_VAR
END_METHOD

END_FUNCTION_BLOCK

// ---- POUs/Prototypes/MeasurementTasks/G6_v_3_5_x/TcoAteqG6_ReadParametersTask_v_3_5_x.TcPOU
(*~
	<docu>
		<summary>
			Read parameters (command bit 5) of the currently selected program: sends Control.ParameterRequest and decodes the response into Status.Parameters. With the map-to-preset flag the list is also mapped onto Status.ParameterSet. Control.QueryParameter is looked up after every read. Read-only - this component never writes parameters.
		</summary>
	</docu>
~*)
FUNCTION_BLOCK TcoAteqG6_ReadParametersTask_v_3_5_x EXTENDS TcoAteqG6Task_v_3_5_x
VAR
	{attribute addProperty Name "<#Map to preset#>"}
	{attribute clr [ReadOnly()]}
	_mapToPreset : BOOL;
END_VAR

IF Execute() THEN
	IF CheckReferences() THEN
		// AX step 0: valid request
		IF _progress = 0 THEN
			inoStatus.ActionDescription := '<#Checking parameter request#>';
			IF TcoAteqG6_IsParameterRequestValid_v_3_5_x(inoRequest := inoControl.ParameterRequest) THEN
				GoTo(10);
			ELSE
				Fail('<#Number of requested parameters out of range (1-35).#>');
			END_IF
		END_IF

		// AX step 10: read and decode
		IF _progress = 10 THEN
			inoStatus.ActionDescription := '<#Reading parameters#>';
			IF Handshake(MASK_READ_PARAMETERS) THEN
				TcoAteqG6_DecodeParameterList_v_3_5_x(inOffset := 16#20,
					inCount := inoControl.ParameterRequest.Count,
					inoImage := inoImage,
					inoList := inoStatus.Parameters);
				IF _mapToPreset THEN
					TcoAteqG6_MapPresetParameters_v_3_5_x(inoList := inoStatus.Parameters, inoSet := inoStatus.ParameterSet);
				END_IF
				TcoAteqG6_QueryParameter_v_3_5_x(inParameter := inoControl.QueryParameter,
					inoList := inoStatus.Parameters,
					inoQuery := inoStatus.ParameterQuery);
				GoTo(100);
			END_IF
		END_IF

		// AX step 100
		IF _progress = 100 THEN
			inoStatus.ActionDescription := '<#Parameters read#>';
			DoneWhen(TRUE);
		END_IF
		Supervise();
	END_IF
END_IF

IF THIS^.Error AND NOT _errorMessage.Pinned THEN
	THIS^.Restore();
END_IF

METHOD FB_init : BOOL
VAR_INPUT
	bInitRetains : BOOL; // if TRUE, the retain variables are initialized (warm start / cold start)
	bInCopyCode : BOOL;  // if TRUE, the instance afterwards gets moved into the copy code (online change)
	ParentObject : ITcoObject;
END_VAR
END_METHOD

METHOD INTERNAL InvokeWithParams : ITcoTaskStatus
VAR_INPUT
	inMapToPreset : BOOL;
END_VAR
IF NOT THIS^.Busy THEN
	_mapToPreset := inMapToPreset;
END_IF
InvokeWithParams := THIS^.Invoke();
END_METHOD

END_FUNCTION_BLOCK
